(* IEC 61131-3 sources: daoli-st-library/DL_Device (part 38) *)

(* ---- FB_DL_AhuDamperStuckDiag.st ---- *)
(*==============================================================================
 * 组件名称 (Component)  : FB_DL_AhuDamperStuckDiag
 * 所属子库 (Sublibrary) : DL_Device
 * 当前版本 (Version)    : 1.0.1
 * 兼容性   (Platform)   : CODESYS 3.5 / TwinCAT 3 / 汇川 InoProShop / Schneider
 *                         Machine Expert；纯 IEC 61131-3（第 3 版）语法，
 *                         仅依赖 Standard.library（R_TRIG / TON）
 * 组件分类 (Category)   : 功能块（FUNCTION_BLOCK）· 设备本体退化诊断 · 风阀卡滞
 * 功能描述 (Function)   : 风阀与电动执行器的卡滞诊断，把含糊的「不动作」拆成
 *                         **三种不同失效机理**——这是本件最大的价值：
 *                         · Full Stall（完全不动）：指令已变、也已得电，但阀位
 *                           **一步未动** → 机械卡死 / 接线断 / 执行器死；
 *                         · Transit Stall（动而未达）：离位了但**没到目标** →
 *                           摩擦力过大 / 气压不足 / 限位错；
 *                         · I/O Fault：反馈信号本身失效 → 传感 / 接线 / 模块
 *                           问题（**不是阀的问题**，误判成阀会导致整台执行器
 *                           被拆下来返修）；
 *                         再加两个工艺级判据：Deviation（稳态偏差超限）与
 *                         Slow（行程时间超标称的设定倍率）。
 * 动作语义 (Semantics)  : 三类失效的处置完全不同：Full Stall 与 I/O Fault 必须
 *                         立刻检修（eFailure）；Transit Stall 亦按 eFailure 处理
 *                         （执行器已失去定位能力）；而 Deviation 与 Slow 是
 *                         **退化**，设备仍可运行（eMaintenanceReq）。三类分开的
 *                         意义就在于此——把「要停机」和「要排计划」分开，而不是
 *                         一个笼统的 bAlarm。
 * 码位级裁定 (Slot rule): `16#0003_0323`（Deviation）落在故障带 `03xx`，但语义是
 *                         「维护请求」，**不置 bError**。理由：bError 表示「不可
 *                         继续运行」，而偏差超限的风阀仍能调节，只是精度不够。
 *                         这是本库首次出现「故障带码 + 不置 bError」的组合，故
 *                         在本头注释显式声明，并要求 MANUAL 故障码表增列
 *                         「是否置 bError」一栏。同理 0161（Slow）为信息级，
 *                         亦不置 bError。`bError` 只由 0321 / 0322 / 0324 / 0325
 *                         四个真正失效的码置位。
 * 段序 (Cycle order)   : 段 1 默认值与单拍预清零 → 段 2 首扫初始化 →
 *                         段 3 参数闸门与输入域判据 → 段 4 定时器与边沿无条件刷新 →
 *                         段 5 复位通道与故障锁存（**CASE 前置，且不做状态赋值**）→
 *                         段 6 状态机 → 段 7 行程与判据累计（含定性）→
 *                         段 8 出口钳位与保持重写 → 段 9 码位链。
 * 定时器清单 (R40)      : 实例名 / IN 表达式 / 断输入拍标志 / 自清位置
 *                         fbTravelWatch / 状态为移动 AND NOT _bTravelBreak
 *                                       / _bTravelBreak（进/出移动态置位）
 *                         fbGraceWatch  / 已超时未达 AND 状态为移动 AND
 *                                       NOT _bTravelBreak / 同上
 *                         fbStallWatch  / 指令已动且阀位未动 AND 状态为移动 AND
 *                                       NOT _bStallBreak / _bStallBreak（进移动态置位）
 *                         fbDevWatch    / 偏差超限 AND 状态为确认 AND
 *                                       NOT _bDevBreak / _bDevBreak（进确认态置位）
 *                         fbSettleWatch / 状态为确认 AND NOT 偏差超限 AND
 *                                       NOT _bSettleBreak / _bSettleBreak（进确认态置位）
 *                         fbIoWatch     / 反馈失效 AND NOT _bIoBreak
 *                                       / _bIoBreak（反馈恢复沿置位）
 *                         六个实例全部在段 4 无条件调用，断输入拍一律在调用后自清。
 * 单拍标志清单 (R25)    : `_bResetPulse` 预清段 1 / 置位段 5 / 消费段 5；
 *                         `_bVerdictPending` 预清段 1 / 置位段 7 / 消费段 7；
 *                         `_bFbRestore` 预清段 1 / 置位段 4 / 消费段 6（恢复首拍）；
 *                         六个断输入标志就地置位、段 4 调用后自清。
 * 保持位清单 (R27)      : `_eDiag`（结论）与 `_fDeviation`、`_tLastTravel`、
 *                         `_uStallCount`、`_uTravelCount` 五个保持量，全部由段 8
 *                         每拍重写出口；复位沿清除。结论在 eVerdict 拍产生后
 *                         **一直保持**，不靠那一个脉冲（R27 正解）。
 * 三元一致表 (R35)      : 量 / 守卫封顶 / 判据运算符
 *                         fSlowRatio   / 钳到 1.1~3.0 / 超时判据用 >=
 *                         fTolPos      / 钳到 0.5~10.0 / 到位判据用 <=
 *                         fDevLimit    / 钳到 1.0~50.0 / 偏差判据用 >
 *                         fDriftThr    / 钳到 0.05~2.0 / 位移判据用 >
 * 验收向量 (Acceptance) :
 *   V1 Full Stall：fCmd 由 0 跳到 60 %、fPosFb 恒 0 → 5 s 后 eDiag=eFullStall、
 *      0321、eHealth=eFailure、bError=TRUE
 *   V2 Transit Stall：fCmd 0→100 %、fPosFb 停在 45 % → 45 s（30 s×1.5）后
 *      但仍在移动则先判 eSlow；若已停止移动则 eTransitStall、0322
 *   V3（V-C 跨段 R40）：连续两次行程（各 20 s 完成，标称 30 s）→ 行程定时器
 *      不得累加到 40 s 判超时；每次进入移动态都必须有断输入拍
 *   V4（V-D 恢复首拍）：bFbValid 由 FALSE 恢复 → 首拍只重装基准，**不判**
 *      Full Stall（否则必误报）
 *   V5（V-A 域外）：fCmd 为 120 % → 钳到 100 并置信息码 0161（钳位不静默）；
 *      fPosFb 为 NaN → 按反馈失效路径处理，且偏差输出夹进 −100~100（R43）
 * 偏离留档 (Deviation)  :
 *   ① 规格 V2 的期望是「45 s 后 eTransitStall」，但 45 s 恰为「1.5 倍标称」的
 *      判据点，此时若阀位仍在缓慢移动，把它判成卡滞会误伤「只是慢」的阀。
 *      本件在 1.5 倍处先置「超时未达」标志，再给一个 tStallTime 的宽限期：
 *      宽限期内到位判 eSlow，超出宽限期仍未到位才判 eTransitStall。这样既
 *      满足 V2 的时序意图，又不把慢阀误判为卡死。
 *   ② 规格未给「确认窗」时长。本件复用 tDevDelay 作为到位确认窗（同一物理
 *      含义：偏差保持在容差内多久算稳定），并在三元一致表登记。
 *   ③ 0161 一码两义：行程慢于 1.5 倍标称，或指令超域被钳位（按 R13 总监
 *      裁定，超域钳位复用该信息码，不新造码位）。
 *   ④ 本件未分到「参数非法」的独立码位，阈值越出物理域（标称行程 <1 s、
 *      倍率越 1.1~3.0、容差或偏差限非正）时复用 0325 兜底码并在本注释登记，
 *      不自行新造码位。
 * 开源溯源 (Origin)     : 来源标签 rockwell-aoi / namur-ne107 / damper-diag。
 *                         原创 clean-room 实现。**仅借鉴 Rockwell AOI（Add-On
 *                         Instruction）公开文档所呈现的「执行器诊断三分类」
 *                         结构粒度**——即把「不动作」拆成完全不动 / 动而未达 /
 *                         反馈失效三类。Rockwell AOI 源码不公开且受其许可协议
 *                         保护，本件**未接触、未复制**任何 AOI 源码、参数名、
 *                         标签名或代码行；三分类的判定阈值、状态机、宽限期
 *                         机制、码位与全部实现细节 100% 本库独立设计。NE107
 *                         （公开推荐规范）仅提供健康分级语义。结构借鉴属功能
 *                         分类层面，不构成代码版权标的，无许可证传染风险。
 * 修订历史 (Revision)   :
 *   2026-11-15  v1.0.0  首版入库（R13 · 泳道 A · 风阀卡滞三分类诊断）
 *   2026-11-16  v1.0.1  终审修复一处（V-C/确认窗类）：判定相的 I/O 失效判据
 *                       由「本拍 NOT _bFbOk」改为「fbIoWatch.Q」，即必须满
 *                       tIoFaultTime 才判 0324；未满时本拍不发布结论、保持上次
 *                       等级。原实现下 eSettling 的到位/偏差定时器（其 IN 不以
 *                       反馈有效性为输入）在反馈刚失效时会无确认窗直接锁存
 *                       0324，属「三分类判据须带确认延时」的缺口。码位与引脚零变化。
 *============================================================================*)

(*-----------------------------------------------------------------------------
 * 枚举: E_DL_DamperDiag（归属本功能块，同文件发布）
 * 含义: 诊断结论。每个成员在段 9 的码位链中有且仅有一个分支，无隐藏成员。
 *-----------------------------------------------------------------------------*)
TYPE E_DL_DamperDiag :
(
    eOk           := 0,    // 正常：无判据成立 / OK, no criterion active
    eSlow         := 10,   // 行程偏慢：超过标称倍率但已到位 / Slow, arrived beyond the ratio
    eDeviation    := 20,   // 稳态偏差：指令与反馈长期不一致 / Steady-state deviation
    eFullStall    := 30,   // 完全卡死：一步未动 / Full stall, not a single step
    eTransitStall := 40,   // 行程卡滞：动了但没到 / Transit stall, moved but never arrived
    eIoFault      := 50    // 反馈失效：信号本身不可信 / Feedback signal lost
);
END_TYPE

(*-----------------------------------------------------------------------------
 * 枚举: E_DL_DamperState（归属本功能块，同文件发布）
 * 含义: 诊断状态机。eMoving 的进出必须与行程定时器挂钩（R40 高危区）。
 *-----------------------------------------------------------------------------*)
TYPE E_DL_DamperState :
(
    eIdle     := 0,    // 待机：偏差在容差内 / Idle, deviation within tolerance
    eMoving   := 10,   // 移动：指令已变且偏差超容差 / Moving, command changed and off target
    eSettling := 20,   // 确认：偏差已进容差，等确认窗 / Settling, waiting for the confirmation window
    eVerdict  := 30,   // 判定：单拍出结论后回待机 / Verdict, single scan then back to idle
    eFault    := 99    // 故障：参数非法或非法状态 / Fault, illegal parameters or state
);
END_TYPE

FUNCTION_BLOCK FB_DL_AhuDamperStuckDiag
VAR_INPUT
    bEnable        : BOOL;                            // 使能 [-] / Enable
    bReset         : BOOL;                            // 复位锁存，上升沿有效 [-] / Rising edge resets the latch
    fCmd           : REAL;                            // 阀位指令 [%]，范围 0~100 / Damper command
    fPosFb         : REAL;                            // 阀位反馈 [%]，范围 0~100 / Position feedback
    bFbValid       : BOOL := TRUE;                    // 反馈有效，AI 断线时为 FALSE [-] / Feedback validity
    bLimitOpen     : BOOL := FALSE;                   // 开到位限位，无此限位时恒 FALSE [-] / Open limit switch
    bLimitClose    : BOOL := FALSE;                   // 关到位限位，无此限位时恒 FALSE [-] / Close limit switch
    tTravelNominal : TIME := T#30S;                   // 全行程标称时间 [毫秒]，范围 1 s~10 min / Nominal full travel time
    fTolPos        : REAL := 3.0;                     // 到位容差 [%]，范围 0.5~10.0 / In-position tolerance
    fDevLimit      : REAL := 10.0;                    // 稳态偏差上限 [%]，范围 1.0~50.0 / Steady-state deviation limit
    tDevDelay      : TIME := T#10S;                   // 偏差确认延时 [毫秒]，范围 0.5~300 s / Deviation confirmation delay
    fDriftThr      : REAL := 0.2;                     // 判有位移的阈值 [%]，范围 0.05~2.0 / Movement threshold
    tStallTime     : TIME := T#5S;                    // 停滞判据时长 [毫秒]，范围 0.5~120 s / Stall duration
    tIoFaultTime   : TIME := T#3S;                    // 反馈失效持续判据 [毫秒]，范围 0.2~60 s / Feedback loss duration
    fSlowRatio     : REAL := 1.5;                     // 判 Slow 的行程倍率 [-]，范围 1.1~3.0 / Slow ratio
END_VAR
VAR_OUTPUT
    eHealth        : E_DL_Ne107Status;                // NE107 健康态（引用自 I_DL_DeviceHealth）[-] / NE107 health
    uDiagCode      : UDINT;                           // 当前诊断码，0=无码 [代码] / Active diagnostic code
    uErrorId       : UDINT;                           // 末次故障码，仅失效级 [代码] / Last fault code
    bError         : BOOL;                            // 故障锁存，仅 0321 0322 0324 0325 置位 [-] / Fault latch
    eDiag          : E_DL_DamperDiag;                 // 诊断结论（保持语义）[-] / Diagnostic verdict, held
    fDeviation     : REAL;                            // 指令减反馈的有符号偏差 [%]，正=开不足 / Signed deviation
    tLastTravel    : TIME;                            // 末次行程实测时间 [毫秒] / Last measured travel time
    nStallCount    : UDINT;                           // 卡滞次数累计 [次]，锁存 / Stall counter
    nTravelCount   : UDINT;                           // 行程次数累计 [次]，锁存 / Travel counter
    bAtOpen        : BOOL;                            // 开到位指示（容差或限位）[-] / At open position
    bAtClose       : BOOL;                            // 关到位指示（容差或限位）[-] / At close position
END_VAR
VAR
    fbTrigReset    : R_TRIG;                          // 复位沿检测，段 4 无条件刷新 [-] / Reset edge detector
    fbFbTrig       : R_TRIG;                          // 反馈恢复沿检测，段 4 无条件刷新 [-] / Feedback restore edge
    fbTravelWatch  : TON;                             // 行程超时计时（标称×倍率），段 4 刷新 [毫秒] / Travel overrun timer
    fbGraceWatch   : TON;                             // 超时后宽限计时，段 4 刷新 [毫秒] / Grace timer after the overrun
    fbStallWatch   : TON;                             // 完全停滞计时，段 4 刷新 [毫秒] / Full stall timer
    fbDevWatch     : TON;                             // 偏差确认计时，段 4 刷新 [毫秒] / Deviation timer
    fbSettleWatch  : TON;                             // 到位确认计时，段 4 刷新 [毫秒] / Settling timer
    fbIoWatch      : TON;                             // 反馈失效计时，段 4 刷新 [毫秒] / Feedback loss timer
    _eState        : E_DL_DamperState := E_DL_DamperState.eIdle; // 当前状态 [-] / Current state
    _bInit         : BOOL := FALSE;                   // 首扫标志，初值 FALSE [-] / First-scan flag
    _bFaultLatch   : BOOL;                            // 故障锁存，仅复位清 [-] / Fault latch
    _uErrFault     : UDINT;                           // 首出故障码 [代码] / First-out fault code
    _uDiagCode     : UDINT;                           // 当前诊断码（单一链产出）[代码] / Active diagnostic code
    _bResetPulse   : BOOL;                            // 复位单拍 [-] / One-shot reset
    _bFbRestore    : BOOL;                            // 反馈恢复单拍 [-] / One-shot restore
    _bVerdictPending : BOOL;                          // 结论待发布单拍 [-] / Verdict pending
    _bTravelBreak  : BOOL;                            // 行程定时器断输入一拍 [-] / Travel timer break
    _bStallBreak   : BOOL;                            // 停滞定时器断输入一拍 [-] / Stall timer break
    _bDevBreak     : BOOL;                            // 偏差定时器断输入一拍 [-] / Deviation timer break
    _bSettleBreak  : BOOL;                            // 确认定时器断输入一拍 [-] / Settling timer break
    _bIoBreak      : BOOL;                            // 反馈失效定时器断输入一拍 [-] / Feedback timer break
    _bOverrun      : BOOL;                            // 行程已超过标称倍率 [-] / Travel overrun flag
    _bCmdOutRange  : BOOL;                            // 指令超域被钳位 [-] / Command clamped flag
    _fCmdUse       : REAL;                            // 生效指令（钳位后）[%] / Effective command
    _fPosUse       : REAL;                            // 生效反馈（钳位后）[%] / Effective position
    _fCmdPrev      : REAL;                            // 上拍指令 [%] / Previous command
    _fPosPrev      : REAL;                            // 上拍反馈 [%] / Previous position
    _fCmdBase      : REAL;                            // 进入移动态的指令基准 [%] / Command baseline at motion start
    _fPosBase      : REAL;                            // 进入移动态的反馈基准 [%] / Position baseline at motion start
    _fTolUse       : REAL := 3.0;                     // 生效到位容差 [%] / Effective tolerance
    _fDevLimitUse  : REAL := 10.0;                    // 生效偏差上限 [%] / Effective deviation limit
    _fDriftUse     : REAL := 0.2;                     // 生效位移阈值 [%] / Effective drift threshold
    _fCmdEpsUse    : REAL := 0.01;                    // 判「指令在动」的极小阈 [%] / Tiny threshold for command motion
    _fSlowUse      : REAL := 1.5;                     // 生效慢速倍率 [-] / Effective slow ratio
    _tTravelUse    : TIME := T#30S;                   // 生效标称行程 [毫秒] / Effective nominal travel
    _tTravelLimit  : TIME := T#45S;                   // 生效超时判据 = 标称×倍率 [毫秒] / Effective travel limit
    _tDevUse       : TIME := T#10S;                   // 生效偏差延时 [毫秒] / Effective deviation delay
    _tStallUse     : TIME := T#5S;                    // 生效停滞时长 [毫秒] / Effective stall duration
    _tIoUse        : TIME := T#3S;                    // 生效反馈失效时长 [毫秒] / Effective feedback loss duration
    _diMs          : DINT;                            // 时间换算中间量 [毫秒] / Time conversion working value
    _fMsReal       : REAL;                            // 行程限值的实数中间量 [毫秒] / Real working value of the travel limit
    _fDeviation    : REAL;                            // 有符号偏差 [%] / Signed deviation
    _bDevExceed    : BOOL;                            // 偏差超限 [-] / Deviation above limit
    _bCmdMovedSince : BOOL;                           // 本行程内指令已动 [-] / Command moved during the travel
    _bPosMovedSince : BOOL;                           // 本行程内阀位已动 [-] / Position moved during the travel
    _bAtTarget     : BOOL;                            // 已到达目标 [-] / Target reached
    _bAtOpenInt    : BOOL;                            // 开到位内部量 [-] / At open internal
    _bAtCloseInt   : BOOL;                            // 关到位内部量 [-] / At close internal
    _bFbOk         : BOOL;                            // 反馈可用（有限且有效）[-] / Feedback usable
    _bFbFinite     : BOOL;                            // 反馈有限标志 [-] / Feedback finite flag
    _bCmdFinite    : BOOL;                            // 指令有限标志 [-] / Command finite flag
    _eDiag         : E_DL_DamperDiag := E_DL_DamperDiag.eOk; // 保持的结论 [-] / Held verdict
    _fDevHeld      : REAL;                            // 保持的偏差 [%] / Held deviation
    _tTravelHeld   : TIME;                            // 保持的末次行程时间 [毫秒] / Held last travel time
    _uStallCount   : UDINT;                           // 保持的卡滞次数 [次] / Held stall counter
    _uTravelCount  : UDINT;                           // 保持的行程次数 [次] / Held travel counter
    _eHealthInt    : E_DL_Ne107Status := E_DL_Ne107Status.eUnknown; // 健康态内部量 [-] / Internal health state
    _bParamBad     : BOOL;                            // 参数非法标志 [-] / Illegal parameter flag
END_VAR
VAR CONSTANT
    DL_VAL_LIM     : REAL := 1.0E6;                   // 有限性判定绝对值上限 [%] / Finiteness limit
    DL_CMD_EPS_RATIO : REAL := 0.05;                  // 指令在动判据相对位移阈的比例 [-] / Command motion ratio
    DL_FULL        : REAL := 100.0;                   // 全行程 [%] / Full stroke
    DL_ZERO        : REAL := 0.0;                     // 零行程 [%] / Zero stroke
    DL_TIME_ZERO   : TIME := T#0S;                    // 时间零值基准 [毫秒] / Time zero reference
    DL_TRAVEL_MIN  : DINT := 1000;                    // 标称行程下限 [毫秒] / Minimum nominal travel
    DL_TRAVEL_MAX  : DINT := 600000;                  // 标称行程上限 [毫秒] / Maximum nominal travel
    DL_DELAY_MIN   : DINT := 500;                     // 延时类下限 [毫秒] / Minimum delay
    DL_DELAY_MAX   : DINT := 300000;                  // 延时类上限 [毫秒] / Maximum delay
    DL_STALL_MIN   : DINT := 500;                     // 停滞时长下限 [毫秒] / Minimum stall duration
    DL_STALL_MAX   : DINT := 120000;                  // 停滞时长上限 [毫秒] / Maximum stall duration
    DL_IO_MIN      : DINT := 200;                     // 反馈失效下限 [毫秒] / Minimum feedback loss
    DL_IO_MAX      : DINT := 60000;                   // 反馈失效上限 [毫秒] / Maximum feedback loss
END_VAR

(*------------------------------------------------------------------------------
 * 段 1｜确定性默认值与单拍标志预清零（R25 第一律）
 *      Deterministic defaults and one-shot flags pre-cleared
 *-----------------------------------------------------------------------------*)
_bResetPulse     := FALSE;                            // 复位单拍预清零（Reset pre-cleared）
_bFbRestore      := FALSE;                            // 恢复单拍预清零（Restore pre-cleared）
_bVerdictPending := FALSE;                            // 结论待发布预清零（Verdict pending pre-cleared）
_bParamBad       := FALSE;                            // 参数非法预清零（Illegal parameter pre-cleared）
_bFbFinite       := FALSE;                            // 反馈有限预清零（Feedback finite pre-cleared）
_bCmdFinite      := FALSE;                            // 指令有限预清零（Command finite pre-cleared）
_bCmdOutRange    := FALSE;                            // 指令超域预清零（Command clamped pre-cleared）

(*------------------------------------------------------------------------------
 * 段 2｜首扫初始化（R19：bInit 初值 FALSE，判据取非；首拍只装基准）
 *      First-scan initialisation, baseline only
 *-----------------------------------------------------------------------------*)
IF NOT _bInit THEN
    _eState       := E_DL_DamperState.eIdle;          // 状态待机（State idle）
    _bFaultLatch  := FALSE;                           // 故障锁存清零（Latch cleared）
    _uErrFault    := 16#0000_0000;                    // 首出码清零（First-out code cleared）
    _eDiag        := E_DL_DamperDiag.eOk;             // 结论正常（Verdict OK）
    _fDevHeld     := 0.0;                             // 偏差保持量清零（Held deviation cleared）
    _tTravelHeld  := DL_TIME_ZERO;                    // 行程时间保持量清零（Held travel cleared）
    _uStallCount  := 0;                               // 卡滞次数清零（Stall counter cleared）
    _uTravelCount := 0;                               // 行程次数清零（Travel counter cleared）
    _fCmdPrev     := 0.0;                             // 上拍指令初值（Previous command）
    _fPosPrev     := 0.0;                             // 上拍反馈初值（Previous position）
    _fCmdBase     := 0.0;                             // 指令基准初值（Command baseline）
    _fPosBase     := 0.0;                             // 反馈基准初值（Position baseline）
    _bOverrun     := FALSE;                           // 超时标志清零（Overrun cleared）
    _bCmdMovedSince := FALSE;                         // 指令位移证据清零（Command evidence cleared）
    _bPosMovedSince := FALSE;                         // 阀位位移证据清零（Position evidence cleared）
    _bInit        := TRUE;                            // 首扫只做一次（First scan runs once）
END_IF

(*------------------------------------------------------------------------------
 * 段 3｜参数闸门、输入域检查与偏差判据（定时器之前，保证本拍值）
 *      Parameter gate, input domain and criteria, ahead of the timers
 *-----------------------------------------------------------------------------*)
_fTolUse      := LIMIT(0.5, fTolPos, 10.0);           // 到位容差钳进 0.5~10 %（Clamped）
_fDevLimitUse := LIMIT(1.0, fDevLimit, 50.0);         // 偏差上限钳进 1~50 %（Clamped）
_fDriftUse    := LIMIT(0.05, fDriftThr, 2.0);         // 位移阈值钳进 0.05~2 %（Clamped）
_fSlowUse     := LIMIT(1.1, fSlowRatio, 3.0);         // 慢速倍率钳进 1.1~3.0（Clamped）
_fCmdEpsUse   := LIMIT(0.001, _fDriftUse * DL_CMD_EPS_RATIO, _fDriftUse); // 指令在动判据，随位移阈缩放并封顶（Scaled and capped）

_diMs        := LIMIT(DL_TRAVEL_MIN, TIME_TO_DINT(tTravelNominal), DL_TRAVEL_MAX); // 标称行程钳位（Clamped）
_tTravelUse  := DINT_TO_TIME(_diMs);                  // 生效标称行程（Effective nominal travel）
_fMsReal     := DINT_TO_REAL(_diMs) * _fSlowUse;      // 超时判据 = 标称 × 倍率 [毫秒]（Limit = nominal times ratio）
_fMsReal     := LIMIT(DINT_TO_REAL(DL_TRAVEL_MIN), _fMsReal, DINT_TO_REAL(DL_TRAVEL_MAX)); // 结果再钳位（Clamped again）
_tTravelLimit := DINT_TO_TIME(REAL_TO_DINT(_fMsReal)); // 生效超时判据（Effective travel limit）

_diMs      := LIMIT(DL_DELAY_MIN, TIME_TO_DINT(tDevDelay), DL_DELAY_MAX); // 偏差延时钳位（Clamped）
_tDevUse   := DINT_TO_TIME(_diMs);                    // 生效偏差延时（Effective deviation delay）
_diMs      := LIMIT(DL_STALL_MIN, TIME_TO_DINT(tStallTime), DL_STALL_MAX); // 停滞时长钳位（Clamped）
_tStallUse := DINT_TO_TIME(_diMs);                    // 生效停滞时长（Effective stall duration）
_diMs      := LIMIT(DL_IO_MIN, TIME_TO_DINT(tIoFaultTime), DL_IO_MAX); // 反馈失效时长钳位（Clamped）
_tIoUse    := DINT_TO_TIME(_diMs);                    // 生效反馈失效时长（Effective feedback loss duration）

(* 输入域检查放在定时器之前：定时器输入要用本拍的可用标志，避免一拍滞后 *)
_bCmdFinite := (fCmd >= -DL_VAL_LIM) AND (fCmd <= DL_VAL_LIM);     // 指令有限（Command finite）
_bFbFinite  := (fPosFb >= -DL_VAL_LIM) AND (fPosFb <= DL_VAL_LIM); // 反馈有限（Feedback finite）
IF (fCmd < DL_ZERO) OR (fCmd > DL_FULL) THEN
    _bCmdOutRange := TRUE;                            // 指令超域：钳位不静默（Clamped, not silent）
END_IF
_fCmdUse := LIMIT(DL_ZERO, fCmd, DL_FULL);            // 指令钳进 0~100 %（Clamped）
IF NOT _bCmdFinite THEN
    _fCmdUse := 0.0;                                  // 非有限：置 0（Non-finite, zeroed）
END_IF
IF _bFbFinite THEN
    _fPosUse := LIMIT(DL_ZERO, fPosFb, DL_FULL);      // 反馈钳进 0~100 %（Clamped）
ELSE
    _fPosUse := _fPosPrev;                            // 非有限：保持上拍值，不污染判据（Hold the previous value）
END_IF
_bFbOk := bFbValid AND _bFbFinite;                    // 反馈可用 = 有效且有限（Usable = valid and finite）

(* 偏差与到位判据：与输入域检查同段，保证定时器用的是本拍值而非上一拍值 *)
_fDeviation  := _fCmdUse - _fPosUse;                  // 有符号偏差，正=开不足（Signed deviation）
_bDevExceed  := _fDeviation > _fDevLimitUse;          // 偏差超限（Deviation above the limit）
_bAtOpenInt  := bLimitOpen OR (_fPosUse >= (DL_FULL - _fTolUse));   // 开到位（At open）
_bAtCloseInt := bLimitClose OR (_fPosUse <= _fTolUse);              // 关到位（At close）
_bAtTarget   := (_fDeviation <= _fTolUse) AND (_fDeviation >= -_fTolUse); // 到位：偏差落在容差带内（In position）

(*------------------------------------------------------------------------------
 * 段 4｜定时器与边沿实例无条件刷新（红线：实例一律在 CASE 之外每拍必调）
 *      Timers and edge detectors refreshed unconditionally outside the CASE
 *-----------------------------------------------------------------------------*)
fbTrigReset(CLK := bReset);                           // 复位沿刷新（Reset edge refreshed）
fbFbTrig(CLK := bFbValid);                            // 反馈恢复沿刷新（Feedback restore edge refreshed）
IF fbFbTrig.Q THEN
    _bFbRestore := TRUE;                              // 反馈恢复单拍（Restore one-shot）
    _bIoBreak   := TRUE;                              // 反馈失效计时重启（Feedback timer restarted）
    _bStallBreak := TRUE;                             // 停滞计时重启，防跨失效期累加（Stall timer restarted）
    _bTravelBreak := TRUE;                            // 行程计时重启（Travel timer restarted）
END_IF

fbTravelWatch(IN := (_eState = E_DL_DamperState.eMoving) AND (NOT _bTravelBreak), PT := _tTravelLimit); // 行程超时计时
(* 宽限计时与行程计时共用同一个断输入拍，故自清必须放在两个实例调用之后，
 * 否则后调的实例永远看不到断输入（R40 的典型陷阱） *)
fbGraceWatch(IN := _bOverrun AND (_eState = E_DL_DamperState.eMoving) AND (NOT _bTravelBreak), PT := _tStallUse); // 宽限计时，断输入沿用行程标志
_bTravelBreak := FALSE;                               // 断输入拍在两个实例调用后自清（Break self-cleared after both calls）

fbStallWatch(IN := _bCmdMovedSince AND (NOT _bPosMovedSince) AND (_eState = E_DL_DamperState.eMoving) AND _bFbOk AND (NOT _bStallBreak), PT := _tStallUse); // 完全停滞计时
_bStallBreak := FALSE;                                // 断输入拍在调用后自清（Break self-cleared）

fbDevWatch(IN := _bDevExceed AND (_eState = E_DL_DamperState.eSettling) AND (NOT _bDevBreak), PT := _tDevUse); // 偏差确认计时
_bDevBreak := FALSE;                                  // 断输入拍在调用后自清（Break self-cleared）

fbSettleWatch(IN := (_eState = E_DL_DamperState.eSettling) AND (NOT _bDevExceed) AND (NOT _bSettleBreak), PT := _tDevUse); // 到位确认计时
_bSettleBreak := FALSE;                               // 断输入拍在调用后自清（Break self-cleared）

fbIoWatch(IN := (NOT _bFbOk) AND (NOT _bIoBreak), PT := _tIoUse); // 反馈失效计时
_bIoBreak := FALSE;                                   // 断输入拍在调用后自清（Break self-cleared)

(*------------------------------------------------------------------------------
 * 段 5｜复位通道 + 故障锁存（CASE 前置；**不做状态变量赋值**，R39）
 *      Reset channel and fault latching before the CASE, with no state write
 *-----------------------------------------------------------------------------*)
IF fbTrigReset.Q THEN
    _bResetPulse := TRUE;                             // 复位单拍（One-shot reset）
END_IF

IF _bResetPulse THEN
    _bFaultLatch  := FALSE;                           // 清故障锁存（Latch cleared）
    _uErrFault    := 16#0000_0000;                    // 清首出码（First-out code cleared）
    _eDiag        := E_DL_DamperDiag.eOk;             // 结论回正常（Verdict back to OK）
    _fDevHeld     := 0.0;                             // 偏差保持量清零（Held deviation cleared）
    _uStallCount  := 0;                               // 卡滞次数清零（Stall counter cleared）
    _uTravelCount := 0;                               // 行程次数清零（Travel counter cleared）
    _bOverrun     := FALSE;                           // 超时标志清零（Overrun cleared）
    _bTravelBreak := TRUE;                            // 行程计时重启（Travel timer restarted）
    _bStallBreak  := TRUE;                            // 停滞计时重启（Stall timer restarted）
    _bDevBreak    := TRUE;                            // 偏差计时重启（Deviation timer restarted）
    _bSettleBreak := TRUE;                            // 确认计时重启（Settling timer restarted）
    _bIoBreak     := TRUE;                            // 反馈计时重启（Feedback timer restarted）
END_IF

(* 参数非法属故障级：行程标称过小会让超时判据恒真，故在闸门处直接判失效 *)
IF (tTravelNominal < T#1S) OR ((fSlowRatio < 1.1) OR (fSlowRatio > 3.0)) THEN
    _bParamBad := TRUE;                               // 参数越出物理域（Parameters outside the physical domain）
END_IF
IF (fTolPos <= 0.0) OR (fDevLimit <= 0.0) THEN
    _bParamBad := TRUE;                               // 容差或偏差限非正（Non-positive tolerance or limit）
END_IF

IF _bParamBad AND (NOT _bFaultLatch) THEN
    _uErrFault   := 16#0003_0325;                     // 0325 非法状态兜底（Illegal configuration fallback）
    _bFaultLatch := TRUE;                             // 锁存（Latched）
END_IF

(*------------------------------------------------------------------------------
 * 段 6｜诊断状态机（5 个成员各一标签 + ELSE 兜底；进出移动态必断行程定时器）
 *      State machine, one label per member plus a trailing fallback
 *-----------------------------------------------------------------------------*)
CASE _eState OF

    E_DL_DamperState.eIdle: // 待机：偏差超容差则按「指令是否变化」分流
        IF _bFaultLatch THEN
            _eState := E_DL_DamperState.eFault;       // 已锁故障（Already latched）
        ELSIF bEnable AND (NOT _bAtTarget) THEN
            IF _bCmdOutRange OR (ABS(_fCmdUse - _fCmdPrev) > _fCmdEpsUse) THEN
                (* 指令已变：进入移动态，装基准并断行程定时器（Command changed, start a travel）
                 * 指令基准取「变化前的上一拍值」，否则基准等于新指令，位移证据永远为假，
                 * 完全停滞判据将永不成立（V1 的核心前提） *)
                _fCmdBase := _fCmdPrev;               // 指令基准取变化前值（Baseline before the change）
                _fPosBase := _fPosUse;                // 反馈基准取当前值（Position baseline）
                _bCmdMovedSince := FALSE;             // 指令位移证据清零（Command evidence cleared）
                _bPosMovedSince := FALSE;             // 阀位位移证据清零（Position evidence cleared）
                _bOverrun := FALSE;                   // 超时标志清零（Overrun cleared）
                _bTravelBreak := TRUE;                // 行程计时断输入一拍后重启（R40）
                _bStallBreak  := TRUE;                // 停滞计时重启（Stall timer restarted）
                IF _uTravelCount < 16#FFFF_FFFF THEN
                    _uTravelCount := _uTravelCount + 1; // 行程次数累加（Travel counter incremented）
                END_IF
                _eState := E_DL_DamperState.eMoving;  // 进入移动态（Enter moving）
            ELSE
                (* 指令未变而偏差超容差：属稳态偏差监视（Steady-state deviation monitoring） *)
                _bDevBreak := TRUE;                   // 偏差计时从 0 起算（Deviation timer restarted）
                _eState := E_DL_DamperState.eSettling; // 进入确认态（Enter settling）
            END_IF
        END_IF

    E_DL_DamperState.eMoving: // 移动：到位则测行程判慢；超时未达判卡滞
        IF _bFaultLatch THEN
            _eState := E_DL_DamperState.eFault;       // 转故障（Enter the fault state）
        ELSIF NOT bEnable THEN
            _bTravelBreak := TRUE;                    // 中止行程计时（Abort the travel timer）
            _eState := E_DL_DamperState.eIdle;        // 回待机（Back to idle）
        ELSIF fbIoWatch.Q THEN
            _bVerdictPending := TRUE;                 // 反馈失效确认（Feedback loss confirmed）
            _bTravelBreak := TRUE;                    // 行程计时中断（Travel timer stopped）
            _eState := E_DL_DamperState.eVerdict;     // 进判定（Enter verdict）
        ELSIF _bFbRestore THEN
            (* 恢复首拍：只重装基准，不判任何卡滞（R41 / V4） *)
            _fCmdBase := _fCmdUse;                    // 重装指令基准（Reload the command baseline）
            _fPosBase := _fPosUse;                    // 重装反馈基准（Reload the position baseline）
            _bCmdMovedSince := FALSE;                 // 位移证据清零（Evidence cleared）
            _bPosMovedSince := FALSE;                 // 位移证据清零（Evidence cleared）
            _bOverrun := FALSE;                       // 超时标志清零（Overrun cleared）
            _bTravelBreak := TRUE;                    // 行程计时重启（Travel timer restarted）
            _bStallBreak := TRUE;                     // 停滞计时重启（Stall timer restarted）
        ELSIF fbStallWatch.Q THEN
            _bVerdictPending := TRUE;                 // 完全停滞确认（Full stall confirmed）
            _bTravelBreak := TRUE;                    // 行程计时中断（Travel timer stopped）
            _eState := E_DL_DamperState.eVerdict;     // 进判定（Enter verdict）
        ELSIF _bAtTarget AND _bFbOk THEN
            _bVerdictPending := TRUE;                 // 到位：出结论（Arrived, issue the verdict）
            _bTravelBreak := TRUE;                    // 行程计时中断（Travel timer stopped）
            _eState := E_DL_DamperState.eVerdict;     // 进判定（Enter verdict）
        ELSIF fbGraceWatch.Q AND _bFbOk THEN
            _bVerdictPending := TRUE;                 // 宽限期满仍未达（Grace expired without arrival）
            _bTravelBreak := TRUE;                    // 行程计时中断（Travel timer stopped）
            _eState := E_DL_DamperState.eVerdict;     // 进判定（Enter verdict）
        END_IF
        (* 反馈暂失时不改状态：保持移动态等内存失效计时，判据由 _bFbOk 抑制 *)

    E_DL_DamperState.eSettling: // 确认：偏差回容差则计确认窗，超限则计偏差窗
        IF _bFaultLatch THEN
            _eState := E_DL_DamperState.eFault;       // 转故障（Enter the fault state）
        ELSIF NOT bEnable THEN
            _bDevBreak := TRUE;                       // 偏差计时中断（Deviation timer stopped）
            _bSettleBreak := TRUE;                    // 确认计时中断（Settling timer stopped）
            _eState := E_DL_DamperState.eIdle;        // 回待机（Back to idle）
        ELSIF _bCmdOutRange OR (ABS(_fCmdUse - _fCmdPrev) > _fCmdEpsUse) THEN
            _bDevBreak := TRUE;                       // 指令又变：回移动态（Command changed again）
            _bSettleBreak := TRUE;                    // 确认计时中断（Settling timer stopped）
            _eState := E_DL_DamperState.eMoving;      // 回移动态（Back to moving）
        ELSIF fbIoWatch.Q THEN
            _bVerdictPending := TRUE;                 // 反馈失效确认（Feedback loss confirmed）
            _eState := E_DL_DamperState.eVerdict;     // 进判定（Enter verdict）
        ELSIF fbDevWatch.Q THEN
            _bVerdictPending := TRUE;                 // 稳态偏差确认（Deviation confirmed）
            _eState := E_DL_DamperState.eVerdict;     // 进判定（Enter verdict）
        ELSIF fbSettleWatch.Q THEN
            _bVerdictPending := TRUE;                 // 确认窗满且无判据（Settled without any criterion）
            _eState := E_DL_DamperState.eVerdict;     // 进判定（Enter verdict）
        END_IF

    E_DL_DamperState.eVerdict: // 判定：结论在段 7 生成，本态只负责回到待机
        _bTravelBreak := TRUE;                        // 出行动态必断行程计时（Leave the motion phase）
        _bStallBreak  := TRUE;                        // 停滞计时重启（Stall timer restarted）
        _bDevBreak    := TRUE;                        // 偏差计时重启（Deviation timer restarted）
        _bSettleBreak := TRUE;                        // 确认计时重启（Settling timer restarted）
        IF _bFaultLatch THEN
            _eState := E_DL_DamperState.eFault;       // 已锁故障优先（Latched fault wins）
        ELSE
            _eState := E_DL_DamperState.eIdle;        // 结论保持，回待机（Verdict held, back to idle）
        END_IF

    E_DL_DamperState.eFault: // 故障：等复位
        IF _bResetPulse THEN
            _eState := E_DL_DamperState.eIdle;        // 复位受理（Reset accepted）
        END_IF

    ELSE
        _uErrFault   := 16#0003_0325;                 // 0325 非法状态兜底（Illegal state fallback）
        _bFaultLatch := TRUE;                         // 兜底锁存（Fallback latched）
        _eState      := E_DL_DamperState.eFault;      // 进终端安全态（Terminal safe state）
END_CASE

(*------------------------------------------------------------------------------
 * 段 7｜行程证据累计与判据定性（在移动/确认/判定三态内推进）
 *      Travel evidence and criterion classification
 *-----------------------------------------------------------------------------*)
IF (_eState = E_DL_DamperState.eMoving) THEN
    IF ABS(_fCmdUse - _fCmdBase) > _fDriftUse THEN
        _bCmdMovedSince := TRUE;                      // 指令已动（Command has moved）
    END_IF
    IF ABS(_fPosUse - _fPosBase) > _fDriftUse THEN
        _bPosMovedSince := TRUE;                      // 阀位已动（Position has moved）
    END_IF
    IF fbTravelWatch.Q THEN
        _bOverrun := TRUE;                            // 超过标称倍率，进入宽限期（Overrun, start the grace window）
    END_IF
END_IF

IF _bVerdictPending THEN
    IF fbIoWatch.Q THEN
        _eDiag := E_DL_DamperDiag.eIoFault;           // 反馈失效满确认窗：不是阀的问题（Feedback fault, not the valve）
        _uErrFault := 16#0003_0324;                   // 0324 I/O 反馈失效（Feedback lost）
        _bFaultLatch := TRUE;                         // 失效级锁存（Failure latch）
    ELSIF NOT _bFbOk THEN
        (* 判定拍反馈失效但未满 tIoFaultTime：本拍**不发布任何结论**，保持上次值。
         * 这是 R42 本拍复验与「三分类判据一律带确认窗」的交点：eSettling 的
         * 到位/偏差定时器不以反馈有效性为输入，若在此直接判 I/O 失效，就会用
         * 一次瞬时断线否掉整段行程；正确路径是让 fbIoWatch 计时满后再定性。 *)
    ELSIF fbStallWatch.Q THEN
        _eDiag := E_DL_DamperDiag.eFullStall;         // 完全不动（Full stall）
        _uErrFault := 16#0003_0321;                   // 0321 Full Stall（Full stall）
        _bFaultLatch := TRUE;                         // 失效级锁存（Failure latch）
        IF _uStallCount < 16#FFFF_FFFF THEN
            _uStallCount := _uStallCount + 1;         // 卡滞计数（Stall counter incremented）
        END_IF
    ELSIF _bAtTarget THEN
        _tTravelHeld := fbTravelWatch.ET;             // 实测行程时间（Measured travel time）
        IF _bOverrun THEN
            _eDiag := E_DL_DamperDiag.eSlow;          // 超时但到位：只是慢（Arrived late, merely slow）
        ELSE
            _eDiag := E_DL_DamperDiag.eOk;            // 准时到位（Arrived in time）
        END_IF
    ELSIF fbGraceWatch.Q THEN
        IF _bPosMovedSince THEN
            _eDiag := E_DL_DamperDiag.eTransitStall;  // 动而未达（Moved but never arrived）
            _uErrFault := 16#0003_0322;               // 0322 Transit Stall（Transit stall）
            _bFaultLatch := TRUE;                     // 失效级锁存（Failure latch）
        ELSE
            _eDiag := E_DL_DamperDiag.eFullStall;     // 一步未动（Not a single step）
            _uErrFault := 16#0003_0321;               // 0321 Full Stall（Full stall）
            _bFaultLatch := TRUE;                     // 失效级锁存（Failure latch）
        END_IF
        IF _uStallCount < 16#FFFF_FFFF THEN
            _uStallCount := _uStallCount + 1;         // 卡滞计数（Stall counter incremented）
        END_IF
    ELSIF fbDevWatch.Q THEN
        _eDiag := E_DL_DamperDiag.eDeviation;         // 稳态偏差：可运行，不置 bError（Deviation, still runnable）
    ELSE
        _eDiag := E_DL_DamperDiag.eOk;                // 无判据（No criterion）
    END_IF
    _bVerdictPending := FALSE;                        // 本拍结论已处理（或按确认窗规则不出结论），标志自清（Verdict consumed）
END_IF

_fDevHeld := LIMIT(-DL_FULL, _fDeviation, DL_FULL);   // 偏差保持量钳进 −100~100（R43）
_fCmdPrev := _fCmdUse;                                // 记录上拍指令（Record the previous command）
_fPosPrev := _fPosUse;                                // 记录上拍反馈（Record the previous position）

(*------------------------------------------------------------------------------
 * 段 8｜健康仲裁、出口钳位与保持重写（R27 + R43）
 *      Health arbitration, clamping and hold semantics
 *-----------------------------------------------------------------------------*)
IF _bFaultLatch THEN
    _eHealthInt := E_DL_Ne107Status.eFailure;         // 失效（Failure）
ELSIF _eDiag = E_DL_DamperDiag.eSlow THEN
    _eHealthInt := E_DL_Ne107Status.eMaintenanceReq;  // 慢：维护请求（Slow, maintenance）
ELSIF _eDiag = E_DL_DamperDiag.eDeviation THEN
    _eHealthInt := E_DL_Ne107Status.eMaintenanceReq;  // 偏差：维护请求（Deviation, maintenance）
ELSIF NOT bEnable THEN
    _eHealthInt := E_DL_Ne107Status.eUnknown;         // 未使能（Disabled）
ELSE
    _eHealthInt := E_DL_Ne107Status.eOk;              // 正常（OK）
END_IF

eHealth      := _eHealthInt;                          // 健康态出口（Health outlet）
eDiag        := _eDiag;                               // 结论保持重写（Held verdict rewritten）
fDeviation   := _fDevHeld;                            // 偏差钳位出口（Clamped deviation）
tLastTravel  := _tTravelHeld;                         // 末次行程时间出口（Last travel outlet）
nStallCount  := _uStallCount;                         // 卡滞次数出口（Stall counter outlet）
nTravelCount := _uTravelCount;                        // 行程次数出口（Travel counter outlet）
bAtOpen      := _bAtOpenInt;                          // 开到位出口（At open outlet）
bAtClose     := _bAtCloseInt;                         // 关到位出口（At close outlet）
bError       := _bFaultLatch;                         // 故障位只由失效级码置位（Failure codes only）

(*------------------------------------------------------------------------------
 * 段 9｜码位单一优先级链（全拍只写一次 uDiagCode）
 *      Single priority chain, the diagnostic code is written exactly once
 *-----------------------------------------------------------------------------*)
IF _bFaultLatch THEN
    _uDiagCode := _uErrFault;                         // 失效级优先（Failure first）
ELSIF _eDiag = E_DL_DamperDiag.eDeviation THEN
    _uDiagCode := 16#0003_0323;                       // 0323 稳态偏差：故障带码但**不置 bError**（Deviation, no bError）
ELSIF (_eDiag = E_DL_DamperDiag.eSlow) OR _bCmdOutRange THEN
    _uDiagCode := 16#0003_0161;                       // 0161 行程偏慢或指令超域钳位（Slow or clamped command）
ELSIF NOT _bFbOk THEN
    _uDiagCode := 16#0003_0160;                       // 0160 无反馈运行，尚未超失效时长（Open-loop run）
ELSE
    _uDiagCode := 16#0000_0000;                       // 无码（No code）
END_IF

uDiagCode := _uDiagCode;                              // 诊断码出口（Diagnostic code outlet）
uErrorId  := _uErrFault;                              // 末次故障码出口（Last fault code outlet）

END_FUNCTION_BLOCK

(* ---- FB_DL_AnalogSensorHealthClassify.st ---- *)
(*==============================================================================
 * 组件名称 (Component)  : FB_DL_AnalogSensorHealthClassify
 * 所属子库 (Sublibrary) : DL_Device ｜ 版本 (Version) : 1.0.2 ｜ 2026-11-23
 * 兼容性   (Platform)   : CODESYS 3.5+ / TwinCAT 3 / 汇川 InoProShop / 施耐德 Machine Expert
 *                         仅依赖 IEC 61131-3 标准（TON / CASE / SQRT 标准函数），零厂商私有库
 * 功能描述 (Function)   : 模拟量通道健康分级（统计窗口径）：在长度 tWinTime 的滑动统计窗内
 *                         累计样本数 / 和 / 平方和 / 最小 / 最大，窗末算出均值 μ 与方差 σ²，
 *                         按四条判据分级：
 *                         · 超量程：本拍样本 > fRangeMax（上侧）或 < fRangeMin（下侧）——即时判，
 *                           上/下各占独立健康成员（R190 归因唯一，禁合并）；
 *                         · 噪声过大：σ² > fNoiseVarMax（窗口级）；
 *                         · 卡滞：σ² < fVarStuckMax 连续 nStuckWinNeed 个统计窗（持续判，
 *                           单窗低方差不算卡滞——慢变工艺量单窗内方差天然很小）；
 *                         · 正常：以上皆否。
 *                         同时输出置信码 nConfidence（0..100），供 HMI 分级显示与预测性维护。
 *                         **与 4-20mA 断线件的分工**：断线 / NE43 电平分级归
 *                         FB_DL_AnalogSignalHealth；本件只看统计特征，不做电平判据。
 * 接口     (Interface)  : 输入 bEnable / bReset / fValue（本拍样本）/ fRangeMin / fRangeMax /
 *                         tWinTime（统计窗长）/ fVarStuckMax / fNoiseVarMax / nStuckWinNeed；
 *                         输出 eHealth（E_DL_AscHealth）/ nConfidence / fMean / fMin / fMax /
 *                         fVar / eState / bError / eCause / bValid。
 * 状态迁移表 (State Transition Table)：
 *   ① eIdle → eCollect：bEnable 上升（开始采样）；拍 N 进入（使能）/ 本拍行为：清统计量、
 *      不判级 / 拍 N+1 转出至 eCollect。
 *   ② eCollect → eClassify：tonWin.Q（统计窗到时）；拍 N 进入（窗到时）/ 本拍行为：
 *      本拍样本不入账（入账发生在 eCollect 拍）/ 拍 N+1 转出至 eClassify。
 *   ③ eClassify → eCollect：分级完成并清统计累加器（同拍完成，单拍驻留）；拍 N 进入 /
 *      本拍行为：算 μ、σ²、判四级、清窗 / 拍 N+1 转出至 eCollect。
 *   ④ eCollect / eClassify → eFault：组态域闸失败（量程倒置 / 窗长 ≤0 / 阈值倒置 /
 *      非有限入参 / nStuckWinNeed < 1）；拍 N 进入（判据失败）/ 本拍行为：锁存首因、
 *      eHealth := eUnknown、nConfidence := 0 / 拍 N+1 转出至 eFault（段尾迁移闸）。
 *   ⑤ eCollect → eIdle：bEnable 落 FALSE（失能退出，健康值冻结为 eUnknown 并置 eNoSample）。
 *   ⑥ eFault → eIdle：bReset 上升且 NOT bEnable（可达性自证 R152：两引脚外部恒可达）；
 *      拍 N 进入 / 本拍行为：清锁存与成因 / 拍 N+1 转出至 eIdle。
 *   ⑦ ELSE（非法枚举值）→ eFault，成因 eIllegalState（R6 兜底）。
 * 边界     (Boundary)   : ① 统计窗 TON 自复位：IN := (状态 = eCollect) AND NOT tonWin.Q
 *                            AND (NOT 故障锁存)（R188 / FB50-1③），不依赖外部沿清零。
 *                         ② 方差公式 σ² = E[x²] − μ²，样本数 n ≥ 1 才计算；n = 0 时置
 *                            信息级 eNoSample 并跳过（除零结构性不可达，R4）。
 *                         ③ 方差可能出现 −1E−18 级负残差（浮点相减），取 MAX(σ², 0) 归零。
 *                         ④ 均值 / 方差 / 极值仅在窗末刷新，窗内保持上一窗结果（不逐拍抖动）。
 *                         ⑤ 浮点同值比较统一容差 DL_ASC_EPS（1E-6），禁 `=`。
 *                         ⑥ 零全局耦合（无 GVL / VAR_EXTERNAL / %I / %Q）。
 * 码表     (Codes)      : 本件不占用全局数字码位（R297 零码位范式）；出口为 BOOL + ENUM，
 *                         enum E_DL_AscCause 归属本文件（全库唯一属主）。信息级
 *                         eNoSample / eWinDone 永不置 bError；故障级码锁存回放至 bReset 沿。
 * 分工声明 (Scope)      : 4-20mA 断线 / NE43 分级归 FB_DL_AnalogSignalHealth；通用信号冻结
 *                         监视归 FB_DL_SignalStuckWatch；窗内中值 / 均值滤波归
 *                         FB_DL_MedianFilter / FB_DL_MovingAverage。
 * 归属     (Ownership)  : E_DL_AscHealth / E_DL_AscPhase / E_DL_AscCause 归属本文件
 *                         （全库唯一定义，R264）；E_DL_AshHealth 属主为
 *                         FB_DL_AnalogSignalHealth.st，本件不引用亦不重声明。
 * 红线自检 (Redline)    : R1 ✓ 零 GVL ｜ R2 ✓ 零 %I/%Q ｜ R3 ✓ 纯 IEC ｜ R4 ✓ 样本数闸防除零 +
 *                         非有限双判 + 容差比较 ｜ R5 ✓ 逐行同行双语注释 ｜ R6 ✓ 三态 ENUM +
 *                         CASE + ELSE ｜ R7 ✓ tonWin 在 CASE 外无条件调用 ｜ R14 ✓ 无 PROPERTY
 *                         R8/R9 N/A（无 METHOD）｜ FB50-1① ✓ CASE 内无 TON 调用
 * 修订历史 (Revision)   : 2026-11-23  v1.0.0  R78-B3 首版
 * 验收向量 (Acceptance) :
 *   V1 量程 0..100、样本恒为 50.0、窗长 1s：首窗 σ²=0 → 第 1 窗不判卡滞（nStuckWinNeed=3），
 *      连续 3 窗后 eHealth=eStuck、nConfidence=20。
 *   V2 样本在 40..60 间交替（σ²≈100）、fNoiseVarMax=10 → eHealth=eNoisy、nConfidence=40。
 *   V3 样本 105.0（> fRangeMax=100）→ 当拍 eHealth=eOverHigh、nConfidence=10（不等窗末）。
 *   V4 fRangeMin=100、fRangeMax=0（倒置）→ eState=eFault、eCause=eBadConfig、bError=TRUE；
 *      bReset 上升且 bEnable=FALSE → 回 eIdle。
 *   V5 tWinTime=T#0s → eState=eFault、eCause=eBadConfig（窗长越域）。
 *============================================================================*)

(*-----------------------------------------------------------------------------
 * 枚举: E_DL_AscHealth（通道健康分级；超量程上/下独立成员，R190）
 *----------------------------------------------------------------------------*)
TYPE E_DL_AscHealth :
(
    eUnknown  := 0,    // 未知：未采样 / 未成窗 / 故障 / Unknown: not sampled or faulted
    eNormal   := 10,   // 正常：窗内方差在带内且未超量程 / Normal: variance in band and within range
    eStuck    := 20,   // 卡滞：连续多窗方差低于阈值 / Stuck: variance below threshold for several windows
    eOverHigh := 30,   // 超量程（上侧）：样本 > fRangeMax / Over range high: sample above the high limit
    eOverLow  := 40,   // 超量程（下侧）：样本 < fRangeMin / Over range low: sample below the low limit
    eNoisy    := 50    // 噪声过大：窗内方差 > fNoiseVarMax / Noisy: window variance above the noise limit
);
END_TYPE

(*-----------------------------------------------------------------------------
 * 枚举: E_DL_AscPhase（状态机相位；eFault 为安全相，仅 bReset 沿迁出）
 *----------------------------------------------------------------------------*)
TYPE E_DL_AscPhase :
(
    eIdle     := 0,    // 空闲：未使能，不采样 / Idle: disabled, no sampling
    eCollect  := 10,   // 采样：逐拍累计统计量 / Collect: accumulate statistics per scan
    eClassify := 20,   // 分级：单拍窗末计算 μ、σ² 并判级 / Classify: single-scan window evaluation
    eFault    := 90    // 故障安全相：组态非法，锁存成因 / Fault safe phase with a latched cause
);
END_TYPE

(*-----------------------------------------------------------------------------
 * 枚举: E_DL_AscCause（成因码；信息级 = 0..9，故障级 = 10 起）
 *----------------------------------------------------------------------------*)
TYPE E_DL_AscCause :
(
    eNone         := 0,   // 信息级：无事件 / Info: no event
    eNoSample     := 1,   // 信息级：窗内无样本（已跳过方差计算）/ Info: no sample in the window, variance skipped
    eWinDone      := 2,   // 信息级：统计窗完成 / Info: statistics window completed
    eBadConfig    := 10,  // 故障级：量程倒置 / 窗长 ≤0 / 阈值倒置 / Fault: inverted range, zero window or inverted thresholds
    eNonFinite    := 11,  // 故障级：入参非有限 / Fault: non-finite input
    eBadWinNeed   := 12,  // 故障级：卡滞窗数需求 < 1 / Fault: stuck window count below one
    eIllegalState := 13   // 故障级：非法状态枚举值 / Fault: illegal state enum value
);
END_TYPE

FUNCTION_BLOCK FB_DL_AnalogSensorHealthClassify
VAR_INPUT
    bEnable      : BOOL := FALSE;      // 使能：FALSE 停止采样（健康值冻结 eUnknown）/ Enable, FALSE stops sampling
    bReset       : BOOL := FALSE;      // 复位（上升沿，需同时 bEnable=FALSE）/ Reset rising edge, requires disabled state
    fValue       : REAL := 0.0;        // 本拍样本值 [工程单位] / Sample value of this scan
    fRangeMin    : REAL := 0.0;        // 量程下限 [工程单位] / Range low limit
    fRangeMax    : REAL := 100.0;      // 量程上限，域 > fRangeMin [工程单位] / Range high limit, domain > fRangeMin
    tWinTime     : TIME := T#1S;       // 统计窗长，域 > 0 [s] / Statistics window length, domain > 0
    fVarStuckMax : REAL := 0.01;       // 卡滞方差阈值（σ² < 该值判疑似卡滞），域 ≥ 0 / Stuck variance threshold, domain >= 0
    fNoiseVarMax : REAL := 25.0;       // 噪声方差阈值（σ² > 该值判噪声过大），域 > fVarStuckMax / Noise variance threshold
    nStuckWinNeed : INT := 3;          // 连续低方差窗数需求，域 ≥ 1 [-] / Consecutive low-variance windows required
END_VAR
VAR_OUTPUT
    eHealth      : E_DL_AscHealth := E_DL_AscHealth.eUnknown;  // 健康分级出口 [-] / Health classification outlet
    nConfidence  : INT := 0;                     // 置信码 0..100（100 = 完全可信）[-] / Confidence code 0..100
    fMean        : REAL := 0.0;                  // 上一窗均值 μ [工程单位] / Mean of the last window
    fMin         : REAL := 0.0;                  // 上一窗最小值 [工程单位] / Minimum of the last window
    fMax         : REAL := 0.0;                  // 上一窗最大值 [工程单位] / Maximum of the last window
    fVar         : REAL := 0.0;                  // 上一窗方差 σ² [(工程单位)²] / Variance of the last window
    eState       : E_DL_AscPhase;                // 状态出口（段尾单点映射）[-] / State outlet mapped at the tail
    bError       : BOOL;                         // 故障锁存标志 [-] / Fault latch flag
    eCause       : E_DL_AscCause;                // 成因码出口（故障期锁存回放）[-] / Cause code outlet
    bValid       : BOOL;                         // 分级结果有效回执 [-] / Health result validity receipt
END_VAR
VAR
    _eState      : E_DL_AscPhase := E_DL_AscPhase.eIdle;      // 内部相位（CASE 唯一写入目标）[-] / Internal phase
    _bFaultLatch : BOOL := FALSE;                             // 故障锁存位（仅 bReset 沿清除）[-] / Fault latch bit
    _eCauseLatch : E_DL_AscCause := E_DL_AscCause.eNone;       // 锁存成因码（FB33-1）[-] / Latched cause code
    _eCauseTmp   : E_DL_AscCause := E_DL_AscCause.eNone;       // 本拍首个成因（未锁存）[-] / First cause of this scan
    _bCfgOk      : BOOL := TRUE;                              // 组态与入参闸通过标志 [-] / Configuration gate flag
    _nCnt        : INT := 0;                                  // 窗内样本数 [个] / Sample count in the current window
    _fSum        : LREAL := 0.0;                              // 窗内样本和 [工程单位] / Sum of samples in the window
    _fSumSq      : LREAL := 0.0;                              // 窗内样本平方和 [(工程单位)²] / Sum of squared samples
    _fWinMin     : REAL := 0.0;                               // 窗内最小值（窗内滚动） / Rolling minimum in the window
    _fWinMax     : REAL := 0.0;                               // 窗内最大值（窗内滚动） / Rolling maximum in the window
    _fMeanCalc   : LREAL := 0.0;                              // 窗末均值中间量 / Mean intermediate at window end
    _fVarCalc    : LREAL := 0.0;                              // 窗末方差中间量 / Variance intermediate at window end
    _nStuckWin   : INT := 0;                                  // 连续低方差窗计数（跨窗保持）/ Consecutive low-variance window counter
    _bOverHigh   : BOOL := FALSE;                             // 本拍上侧超量程标志 [-] / Over-range high flag of this scan
    _bOverLow    : BOOL := FALSE;                             // 本拍下侧超量程标志 [-] / Over-range low flag of this scan
    tonWin       : TON;                                       // 统计窗定时器（段 2 无条件调用）/ Statistics window timer, called unconditionally
    _rtReset     : R_TRIG;                                 // 复位沿检测实例（v1.0.2 补：声明沿即实现沿，CASE 外无条件刷新）/ Reset edge detector refreshed outside the CASE
END_VAR
VAR CONSTANT
    DL_ASC_ZERO  : REAL := 0.0;      // 零基准 [-] / Zero base
    DL_ASC_ONE   : REAL := 1.0;      // 一基准（样本数换算用）[-] / Unity base
    DL_ASC_FULL  : REAL := 100.0;    // 置信码满值 [-] / Full confidence value
    DL_ASC_EPS   : REAL := 1.0E-6;   // 浮点同值比较容差 [-] / Float equality tolerance
END_VAR

(* —— 段 1：当拍工作量预置（单拍标志与中间量，不清锁存/累加器/计数） —— *)
_bCfgOk    := TRUE;                                    // 闸通过标志复位 / Gate flag reset
_eCauseTmp := E_DL_AscCause.eNone;                      // 当拍成因复位 / Scan cause reset
_bOverHigh := FALSE;                                    // 上超量程标志复位 / Over-high flag reset
_bOverLow  := FALSE;                                    // 下超量程标志复位 / Over-low flag reset

(* —— 段 2：组态与入参域闸（R272 全量枚举所有浮点与时间引脚） —— *)
IF (fValue <> fValue) OR ((fValue - fValue) <> DL_ASC_ZERO)
    OR (fRangeMin <> fRangeMin) OR ((fRangeMin - fRangeMin) <> DL_ASC_ZERO)
    OR (fRangeMax <> fRangeMax) OR ((fRangeMax - fRangeMax) <> DL_ASC_ZERO)
    OR (fVarStuckMax <> fVarStuckMax) OR ((fVarStuckMax - fVarStuckMax) <> DL_ASC_ZERO)
    OR (fNoiseVarMax <> fNoiseVarMax) OR ((fNoiseVarMax - fNoiseVarMax) <> DL_ASC_ZERO) THEN
    _bCfgOk    := FALSE;
    _eCauseTmp := E_DL_AscCause.eNonFinite;             // 故障级：非有限入参 / Fault: non-finite input
END_IF
IF _bCfgOk THEN
    IF fRangeMax <= fRangeMin THEN
        _bCfgOk    := FALSE;
        _eCauseTmp := E_DL_AscCause.eBadConfig;          // 故障级：量程倒置 / Fault: inverted range
    ELSIF tWinTime <= T#0S THEN
        _bCfgOk    := FALSE;
        _eCauseTmp := E_DL_AscCause.eBadConfig;          // 故障级：窗长越域 / Fault: window length out of domain
    ELSIF fVarStuckMax < DL_ASC_ZERO THEN
        _bCfgOk    := FALSE;
        _eCauseTmp := E_DL_AscCause.eBadConfig;          // 故障级：卡滞阈值为负 / Fault: negative stuck threshold
    ELSIF fNoiseVarMax <= fVarStuckMax THEN
        _bCfgOk    := FALSE;
        _eCauseTmp := E_DL_AscCause.eBadConfig;          // 故障级：噪声阈值不高于卡滞阈值 / Fault: noise threshold not above the stuck one
    ELSIF nStuckWinNeed < 1 THEN
        _bCfgOk    := FALSE;
        _eCauseTmp := E_DL_AscCause.eBadWinNeed;         // 故障级：窗数需求越域 / Fault: window count out of domain
    END_IF
END_IF

(* —— 段 3：统计窗定时器（CASE 外无条件调用；IN 自复位 + 串故障锁存，R188 / FB50-1③） —— *)
tonWin(IN := (_eState = E_DL_AscPhase.eCollect) AND (NOT tonWin.Q) AND (NOT _bFaultLatch),
       PT := tWinTime);                                  // 窗长取引脚（TIME 类型原样传入）/ Window length from the pin

(* —— 段 4：状态机主体（唯一相位写入点） —— *)
_rtReset(CLK := bReset);                                // 复位沿刷新无条件周期调用（R7；v1.0.2 修复 J1 电平判据缺陷 / R18）/ Refresh the reset edge unconditionally every scan
CASE _eState OF
    E_DL_AscPhase.eIdle :
        IF bEnable AND _bCfgOk THEN
            _nCnt      := 0;                             // 清样本计数 / Clear the sample count
            _fSum      := 0.0;                           // 清样本和 / Clear the sum
            _fSumSq    := 0.0;                           // 清平方和 / Clear the squared sum
            _nStuckWin := 0;                             // 清卡滞窗计数 / Clear the stuck window counter
            eHealth    := E_DL_AscHealth.eUnknown;       // 未成窗 → 未知 / Not yet windowed: unknown
            nConfidence := 0;                            // 置信码清零 / Confidence zeroed
            _eState    := E_DL_AscPhase.eCollect;        // 迁移①：进入采样相 / Move to collect
        END_IF

    E_DL_AscPhase.eCollect :
        IF NOT bEnable THEN
            eHealth     := E_DL_AscHealth.eUnknown;      // 迁移⑤：失能后健康值不再成立 / Health no longer valid after disable
            nConfidence := 0;                            // 置信码清零 / Confidence zeroed
            eCause      := E_DL_AscCause.eNoSample;      // 信息级：停止采样 / Info: sampling stopped
            _nStuckWin  := 0;                            // 停采清卡滞计数 / Clear the stuck counter while stopped
            _eState     := E_DL_AscPhase.eIdle;          // 回空闲相 / Back to idle
        ELSE
            (* 逐拍入账（样本数 / 和 / 平方和 / 极值），极值用窗内滚动 *)
            IF _nCnt = 0 THEN
                _fWinMin := fValue;                      // 首样本初始化最小值 / First sample initialises the minimum
                _fWinMax := fValue;                      // 首样本初始化最大值 / First sample initialises the maximum
            ELSE
                _fWinMin := MIN(_fWinMin, fValue);       // 滚动最小 / Rolling minimum
                _fWinMax := MAX(_fWinMax, fValue);       // 滚动最大 / Rolling maximum
            END_IF
            _nCnt   := _nCnt + 1;                        // 样本计数递增 / Increment the sample count
            _fSum   := _fSum + fValue;                   // 累加样本和 / Accumulate the sum
            _fSumSq := _fSumSq + (fValue * fValue);      // 累加平方和 / Accumulate the squared sum
            (* 超量程即时判（上 / 下分列，R146 / R190） *)
            IF fValue > (fRangeMax + DL_ASC_EPS) THEN
                _bOverHigh  := TRUE;                     // 上侧超量程 / Over range high
                eHealth     := E_DL_AscHealth.eOverHigh; // 健康分级立即上报 / Health reported immediately
                nConfidence := 10;                       // 低置信 / Low confidence
                eCause      := E_DL_AscCause.eNone;      // 成因码由健康枚举承担 / Cause expressed by the health enum
            ELSIF fValue < (fRangeMin - DL_ASC_EPS) THEN
                _bOverLow   := TRUE;                     // 下侧超量程 / Over range low
                eHealth     := E_DL_AscHealth.eOverLow;  // 健康分级立即上报 / Health reported immediately
                nConfidence := 10;                       // 低置信 / Low confidence
                eCause      := E_DL_AscCause.eNone;      // 成因码由健康枚举承担 / Cause expressed by the health enum
            END_IF
            IF tonWin.Q THEN
                _eState := E_DL_AscPhase.eClassify;      // 迁移②：窗到时进入分级相 / Window elapsed: move to classify
            END_IF
        END_IF

    E_DL_AscPhase.eClassify :
        IF _nCnt < 1 THEN
            eCause := E_DL_AscCause.eNoSample;           // 信息级：窗内无样本 / Info: no sample in the window
            fMean  := DL_ASC_ZERO;                       // 均值置零哨兵 / Mean sentinel
            fVar   := DL_ASC_ZERO;                       // 方差置零哨兵 / Variance sentinel
            fMin   := DL_ASC_ZERO;                       // 最小值置零哨兵 / Minimum sentinel
            fMax   := DL_ASC_ZERO;                       // 最大值置零哨兵 / Maximum sentinel
            eHealth     := E_DL_AscHealth.eUnknown;      // 分级未知 / Unknown classification
            nConfidence := 0;                            // 置信码清零 / Confidence zeroed
        ELSE
            (* 窗末统计：μ = Σx/n，σ² = Σx²/n − μ²（n ≥ 1，除零不可达） *)
            _fMeanCalc := _fSum / INT_TO_LREAL(_nCnt);                     // 均值 / Mean
            _fVarCalc  := (_fSumSq / INT_TO_LREAL(_nCnt)) - (_fMeanCalc * _fMeanCalc);   // 方差 / Variance
            IF _fVarCalc < 0.0 THEN
                _fVarCalc := 0.0;                                          // 负残差归零（浮点相减残差）/ Negative residual zeroed
            END_IF
            fMean := LREAL_TO_REAL(_fMeanCalc);                            // 均值出口（显式窄化）/ Mean outlet, explicit narrowing
            fVar  := LREAL_TO_REAL(_fVarCalc);                             // 方差出口（显式窄化）/ Variance outlet, explicit narrowing
            fMin  := _fWinMin;                                             // 最小值出口 / Minimum outlet
            fMax  := _fWinMax;                                             // 最大值出口 / Maximum outlet
            eCause := E_DL_AscCause.eWinDone;                              // 信息级：窗完成 / Info: window completed
            (* v1.0.2 补（闸 P1）：_bOverHigh/_bOverLow 段 1 每拍被清，逐拍置位到 eClassify 已不可见
               → 改由窗极值重算，超量程判据真正生效（窗级口径，与头注窗末分级一致） *)
            IF _fWinMax > fRangeMax THEN                                  // 窗内最高样本越上限 / window max above the range
                _bOverHigh := TRUE;                                        // 上超量程成立 / Over-high confirmed
            END_IF
            IF _fWinMin < fRangeMin THEN                                  // 窗内最低样本越下限 / window min below the range
                _bOverLow := TRUE;                                         // 下超量程成立 / Over-low confirmed
            END_IF
            (* 分级：超量程优先（安全侧），其次噪声，再次卡滞，最后正常 *)
            IF _bOverHigh THEN
                eHealth     := E_DL_AscHealth.eOverHigh;                   // 超量程（上）/ Over range high
                nConfidence := 10;                                         // 低置信 / Low confidence
                _nStuckWin  := 0;                                          // 清卡滞计数 / Clear the stuck counter
            ELSIF _bOverLow THEN
                eHealth     := E_DL_AscHealth.eOverLow;                    // 超量程（下）/ Over range low
                nConfidence := 10;                                         // 低置信 / Low confidence
                _nStuckWin  := 0;                                          // 清卡滞计数 / Clear the stuck counter
            ELSIF fVar > fNoiseVarMax THEN
                eHealth     := E_DL_AscHealth.eNoisy;                      // 噪声过大 / Noisy
                nConfidence := 40;                                         // 中低置信 / Medium-low confidence
                _nStuckWin  := 0;                                          // 清卡滞计数 / Clear the stuck counter
            ELSIF fVar < fVarStuckMax THEN
                _nStuckWin := _nStuckWin + 1;                              // 连续低方差窗计数 / Consecutive low-variance windows
                IF _nStuckWin >= nStuckWinNeed THEN
                    eHealth     := E_DL_AscHealth.eStuck;                  // 卡滞（持续判已满足）/ Stuck after the required windows
                    nConfidence := 20;                                     // 低置信 / Low confidence
                ELSE
                    eHealth     := E_DL_AscHealth.eNormal;                 // 尚未满足持续条件：按正常上报 / Not yet persistent: normal
                    nConfidence := 70;                                     // 中等置信 / Medium confidence
                END_IF
            ELSE
                eHealth     := E_DL_AscHealth.eNormal;                     // 正常 / Normal
                nConfidence := 100;                                        // 满置信 / Full confidence
                _nStuckWin  := 0;                                          // 清卡滞计数 / Clear the stuck counter
            END_IF
        END_IF
        (* 清窗（样本数 / 和 / 平方和），极值在下一窗首样本重初始化 *)
        _nCnt   := 0;                                                      // 清样本计数 / Clear the sample count
        _fSum   := 0.0;                                                    // 清和 / Clear the sum
        _fSumSq := 0.0;                                                    // 清平方和 / Clear the squared sum
        _bOverHigh := FALSE;                                               // 清上超量程（窗级标志随窗清零）/ Clear the over-high window flag
        _bOverLow  := FALSE;                                               // 清下超量程 / Clear the over-low window flag
        _eState := E_DL_AscPhase.eCollect;                                 // 迁移③：回到采样相 / Back to collect

    E_DL_AscPhase.eFault :
        (* 迁移⑥：唯一出口 —— bReset 沿 + 已失能 *)
        IF _rtReset.Q AND (NOT bEnable) THEN
            _bFaultLatch := FALSE;                                        // 清故障锁存 / Clear the latch
            _eCauseLatch := E_DL_AscCause.eNone;                          // 清锁存成因 / Clear the latched cause
            eCause       := E_DL_AscCause.eNone;                          // 出口同步 / Outlet follows
            _eState      := E_DL_AscPhase.eIdle;                          // 回空闲相 / Back to idle
        END_IF

ELSE
    (* 迁移⑦：非法枚举兜底（R6） *)
    _eCauseLatch := E_DL_AscCause.eIllegalState;                          // 故障级：非法状态
    _bFaultLatch := TRUE;                                                 // 置锁存 / Latch
    eHealth      := E_DL_AscHealth.eUnknown;                              // 分级未知 / Unknown health
    nConfidence  := 0;                                                    // 置信清零 / Confidence zeroed
    _eState      := E_DL_AscPhase.eFault;                                 // 迁入故障相 / Move to fault
END_CASE

(* —— 段 5：组态闸失败处理（在状态机之后统一置故障，避免分支内重复） —— *)
IF (NOT _bCfgOk) AND (NOT _bFaultLatch) THEN
    _eCauseLatch := _eCauseTmp;                                           // 锁存首因 / Latch the first cause
    _bFaultLatch := TRUE;                                                 // 置故障锁存 / Latch the fault
    eHealth      := E_DL_AscHealth.eUnknown;                              // 分级未知 / Unknown health
    nConfidence  := 0;                                                    // 置信清零 / Confidence zeroed
END_IF

(* —— 段 6：段尾故障迁移闸（锁存与迁相分离，FB50-1④） —— *)
IF _bFaultLatch AND (_eState <> E_DL_AscPhase.eFault) THEN
    _eState := E_DL_AscPhase.eFault;                                       // 锁存即迁相 / Latch forces the fault phase
END_IF

(* —— 段 7：统一出口（状态映射 + 锁存回放） —— *)
eState := _eState;                                                        // 相位映射 / Phase mapping
bError := _bFaultLatch;                                                   // 故障标志取锁存位 / Fault flag from the latch
IF _bFaultLatch THEN
    eCause := _eCauseLatch;                                               // 故障期回放锁存码（FB33-1）/ Replay the latched code
END_IF
bValid := (_eState = E_DL_AscPhase.eCollect) AND (NOT _bFaultLatch) AND (_nCnt > 0);   // 采样相且有样本时有效
END_FUNCTION_BLOCK

(* ---- FB_DL_GuardLockDoor.st ---- *)
(*==============================================================================
 * 组件名称 (Component)  : FB_DL_GuardLockDoor
 * 所属子库 (Sublibrary) : DL_Device
 * 当前版本 (Version)    : 1.0.0
 * 兼容性   (Platform)   : CODESYS 3.5 / TwinCAT 3 / 汇川 InoProShop / Machine Expert
 *                         仅依赖 Standard.library（TON / R_TRIG），零厂商方言
 * 分类     (Category)   : 设备功能块（Function Block，实现 I_DL_SafetyDoor）
 * 功能简述 (Function)   : 带电磁锁扣安全门联锁控制器。时序骨架（ISO 14119
 *                         公开语义 clean-room）：请求解锁 → 停机请求输出 →
 *                         静止确认（零速反馈或 run-down 计时器二选一）→ 解
 *                         锁输出 → 开门审计 → 关门再锁定确认窗 → 复位后才
 *                         允许重启（禁止自动重启）；防篡改冲突诊断、解锁电
 *                         磁铁出口断言式硬约束。
 * 定位声明 (Positioning): 公约 0.13——本块为标准 PLC 逻辑编排与诊断镜像层，
 *                         不构成 ISO 13849 / IEC 62061 认证安全功能，安全回
 *                         路由认证安全控制器/安全 PLC 承载；硬限位与安全门
 *                         开关的最终防线在认证安全回路。
 * 接口实现 (Implements) : I_DL_SafetyDoor。接口属性同名成员（eState/bClosed/
 *                         bLocked/bUnlockPermitted/bOpened/bFault/uErrorId）
 *                         按 R22 以只读 PROPERTY GET 承载（内部镜像同源），
 *                         非接口成员 bUnlockCoil/bStopRequest/uOpenCount 保
 *                         留 VAR_OUTPUT；方法 CmdRequestUnlock/CmdRelock/
 *                         CmdReset/CmdAuditClear 在本文件尾部落地。
 * 公约遵循 (Convention) : 0.1/R23 事件型时序状态机（指令沿 + 反馈电平驱动），
 *                         免首扫，无 bInit。
 *                         0.2/R21 bFault 显式排除信息级码；0.5/R7 全部实例主
 *                         体最前部无条件刷新；0.7/R15 故障级锁存仅复位路径
 *                         清码。
 *                         0.8 故障码段位 16#0003_xxxx（经 DL_Device
 *                         VERSION.md 码表核对：规格建议 0003_0260/0261/0262
 *                         已被 FB_DL_AnalogValve 占用、0003_0105 终审空置，
 *                         依公约冲突顺延）：
 *                         【故障级】0003_0290 静止确认超时（解锁链未达成）、
 *                         0003_0291 门锁不合理组合（防篡改冲突）、0003_0292
 *                         再锁定超时、0003_0293 非法状态兜底；
 *                         【信息级】0003_0121 run-down 计时器模式提示（非零
 *                         速实测，解锁时序期间每拍提示）。
 * 红线自检 (Redline)    : R1 零全局变量表/外部变量引用 ✓｜R2 零物理 IO 地址 ✓
 *                         R3 纯 IEC 61131-3 ✓｜R4 时序超窗防御/出口断言 ✓
 *                         R5 全变量中英双语同行注释 ✓｜R6 ENUM+CASE+ELSE ✓
 *                         R7 五实例（R_TRIG×2/TON×3）主体最前部无条件刷新 ✓
 *                         R8 全常量化 ✓
 * 设计要点 (Key notes)  : ① 解锁链硬约束（出口断言式）：bUnlockCoil 置位前
 *                           提 = （bStandstill 或 tRunDown 计满）AND
 *                           bDoorClosed AND bLockEngaged；三条件不满足时解
 *                           锁输出恒断；
 *                         ② 防篡改冲突：门开（bDoorClosed=FALSE）+ 锁闭反
 *                           馈（bLockEngaged=TRUE）同时为真 → 故障锁存（全
 *                           局监视，任意态生效）；
 *                         ③ 关门再锁定：关门沿 → 锁闭反馈确认窗（常量
 *                           DL_RELOCK_WINDOW）内未闭 → 故障；
 *                         ④ 重启抑制：开门事件后必须 bReset 且门锁全确认才
 *                           回 eIdle，无任何自动重启路径；
 *                         ⑤ tRunDown 按实测最差停机时间整定，制动维护后必
 *                           须重测（引脚注释与手册口径）。
 * 偏离留档 (Deviation)  : 依 R11 头注释留档，共 1 条：
 *                         ① 码位顺延：规格建议 0003_0260/0261/0262 与既有
 *                           FB_DL_AnalogValve 冲突、0003_0105 空置，依公约
 *                           0.8 顺延为 0003_0290/0291/0292/0293 与
 *                           0003_0121（核对结果优先于建议值）。
 * 开源溯源 (Origin)     : 来源标签 tcopen-component / safety-interlock
 *                         （RAW_NOTES_R7 S-4：ISO 14119 电磁锁扣门联锁公开
 *                         语义——解锁时序骨架、run-down 计时、防篡改诊断，
 *                         公开标准资料，仅借鉴语义域；状态机、出口断言、码
 *                         位与引脚契约 100% 本库独立设计，clean-room 未复
 *                         制源码）。
 * 验收向量 (Acceptance) :
 *   V1 解锁全链（零速模式）：请求 → eStopRequested → bStandstill=TRUE →
 *      eStandstillConfirmed → eUnlocked → 开门 → eOpened 审计+1；
 *   V2 run-down 模式计时链：bUseStandstillFb=FALSE → tRunDown 计满 → 解锁，
 *      期间信息级 0003_0121；
 *   V3 静止确认超时：eStopRequested 超 DL_UNLOCK_TIMEOUT → 故障 0003_0290；
 *   V4 防篡改冲突注入：门开+锁闭反馈同真 → 故障 0003_0291（任意态生效）；
 *   V5 开门审计与再锁定：关门沿 → DL_RELOCK_WINDOW 内锁闭确认 → eLocked；
 *      超窗 → 0003_0292；
 *   V6 复位后重启抑制：再锁定完成 + bReset 沿 → eIdle；无 bReset 时解锁请
 *      求被拒（bUnlockPermitted=FALSE）。
 * 修订历史 (Revision)   :
 *   2026-11-15  v1.0.0  首版入库（Round 07 · DL_Device 安全门族实现件）
 *============================================================================*)
FUNCTION_BLOCK FB_DL_GuardLockDoor IMPLEMENTS I_DL_SafetyDoor
VAR_INPUT
    bCmdUnlock       : BOOL;            // 解锁请求指令（Unlock request），上升沿发起解锁时序 / Unlock request edge starts the sequence
    bCmdRelock       : BOOL;            // 重新闭锁指令（Relock command），电平生效 / Relock command, level effective
    bReset           : BOOL;            // 上升沿复位故障与重启抑制（Reset edge clears fault and restart inhibit）/ Reset edge
    bDoorClosed      : BOOL;            // 门关闭反馈（Door closed feedback），TRUE=门已关；NC 语义由接线层保证 / Door closed, NC semantics by wiring layer
    bLockEngaged     : BOOL;            // 锁闭反馈（Lock engaged feedback），TRUE=机械锁扣已闭 / Lock engaged, TRUE = mechanical lock closed
    bStandstill      : BOOL;            // 静止确认反馈（Standstill feedback，可选零速信号），TRUE=危险运动已停止 / Standstill feedback, TRUE = hazardous motion stopped
    bUseStandstillFb : BOOL;            // 静止反馈使能（Standstill feedback enable），TRUE=用 bStandstill 判静止；FALSE=用 run-down 计时器 / TRUE = zero-speed mode, FALSE = run-down timer mode
    tRunDown         : TIME := T#5S;    // 停机走完计时（Run-down time），默认 T#5S；按实测最差停机时间整定，制动维护后重测 / Run-down time, tune to measured worst-case stopping time, re-measure after brake maintenance
END_VAR
VAR_OUTPUT
    bUnlockCoil : BOOL;                 // 解锁电磁铁输出（Unlock solenoid coil），断电解锁方向（失电=保持锁定，弹簧锁语义）/ Unlock coil, de-energize-to-unlock (spring-lock semantics)
    bStopRequest: BOOL;                 // 停机请求输出（Stop request），解锁时序中置位直到静止确认 / Stop request active during the unlock sequence until standstill confirmed
    uOpenCount  : UDINT;                // 开门次数审计（Open audit count），CmdAuditClear 清零 / Open audit count, cleared by CmdAuditClear
END_VAR
VAR
    _eState         : E_DL_SafetyDoorState := E_DL_SafetyDoorState.eIdle; // 内部时序状态（Internal sequence state），属性只读 / Internal state, read-only via property
    _bFaultLatch    : BOOL;            // 故障锁存标志（Fault latch flag），仅复位路径清除 / Fault latch, cleared only via reset path
    _uErrorIdInt    : UDINT;           // 内部故障级码寄存（Internal fault-level register）/ Internal fault-level register
    _uInfoCode      : UDINT;           // 本拍信息级码（Info code this cycle），瞬时型每拍重算 / Transient info code, recomputed each scan
    _bRestartInhibit: BOOL;            // 重启抑制标志（Restart inhibit），开门事件置位、复位沿清除 / Restart inhibit, set on open event, cleared by reset
    _bRelockCheck   : BOOL;            // 再锁定确认窗计时中（Relock confirm window running）/ Relock confirm window running
    _bPendUnlock    : BOOL;            // 方法解锁请求（Method unlock request）/ Method unlock request
    _bPendRelock    : BOOL;            // 方法再闭锁请求（Method relock request）/ Method relock request
    _bPendReset     : BOOL;            // 方法复位请求（Method reset request）/ Method reset request
    _bPendAuditClr  : BOOL;            // 方法审计清除请求（Method audit-clear request）/ Method audit-clear request
    _bUnlockReq     : BOOL;            // 合成解锁请求（Merged unlock request），引脚沿 OR 方法 / Merged unlock request
    _bStandstillOk  : BOOL;            // 静止确认达成（Standstill achieved），零速反馈或计时器二选一 / Standstill achieved by either source
    _fbTrigUnlock   : R_TRIG;          // 解锁请求沿（Unlock request edge）/ Unlock request edge detector
    _fbTrigReset    : R_TRIG;          // 复位沿（Reset edge）/ Reset edge detector
    _fbTonRunDown   : TON;             // run-down 计时器（Run-down timer），计时器模式判静止 / Run-down timer for timer-mode standstill
    _fbTonUnlockTo  : TON;             // 解锁链超时监视（Unlock-chain timeout monitor）/ Unlock-chain timeout monitor
    _fbTonRelockWin : TON;             // 再锁定确认窗（Relock confirm window）/ Relock confirm window
END_VAR
VAR CONSTANT
    DL_RELOCK_WINDOW  : TIME := T#2S;   // 再锁定确认窗（Relock confirm window），窗内未闭锁即故障 / Relock confirm window, no engagement in window = fault
    DL_UNLOCK_TIMEOUT : TIME := T#30S;  // 解锁链总超时（Unlock-chain timeout），静止确认未达即故障 / Unlock-chain timeout for standstill confirmation
END_VAR

METHOD CmdRequestUnlock : BOOL
VAR_INPUT
END_VAR
IF _bFaultLatch OR (_eState = E_DL_SafetyDoorState.eFault) OR (NOT bDoorClosed) THEN
    CmdRequestUnlock := FALSE;    // 故障态/门开态拒绝（Rejected in fault or door-open）
ELSE
    _bPendUnlock := TRUE;         // 登记解锁请求，主体状态机消化（Register unlock, consumed by body）
    CmdRequestUnlock := TRUE;     // 受理成功（Accepted）
END_IF

(*------------------------------------------------------------------------------
 * 方法: CmdRelock —— 重新闭锁指令：门开态下关门后受理。
 *      Method CmdRelock - relock, accepted on door close in opened state.
 *------------------------------------------------------------------------------*)
    END_METHOD

METHOD CmdRelock : BOOL
VAR_INPUT
END_VAR
IF (_eState = E_DL_SafetyDoorState.eOpened) AND bDoorClosed THEN
    _bPendRelock := TRUE;         // 登记再闭锁请求（Register relock request）
    CmdRelock := TRUE;            // 受理成功（Accepted）
ELSE
    CmdRelock := FALSE;           // 非门开态/门未关拒绝（Rejected outside opened-with-closed-door）
END_IF

(*------------------------------------------------------------------------------
 * 方法: CmdReset —— 复位故障：仅故障态受理（接口方法拒绝语义红线）。
 *      Method CmdReset - reset, accepted only in fault state.
 *------------------------------------------------------------------------------*)
    END_METHOD

METHOD CmdReset : BOOL
VAR_INPUT
END_VAR
IF _bFaultLatch OR (_eState = E_DL_SafetyDoorState.eFault) THEN
    _bPendReset := TRUE;          // 登记复位请求（Register reset request）
    CmdReset := TRUE;             // 可复位（Resettable）
ELSE
    CmdReset := FALSE;            // 无故障可复位（Nothing to reset）
END_IF

(*------------------------------------------------------------------------------
 * 方法: CmdAuditClear —— 清除开门审计记录：故障态拒绝。
 *      Method CmdAuditClear - clears the open audit count, rejected in fault.
 *------------------------------------------------------------------------------*)
    END_METHOD

METHOD CmdAuditClear : BOOL
VAR_INPUT
END_VAR
IF _bFaultLatch OR (_eState = E_DL_SafetyDoorState.eFault) THEN
    CmdAuditClear := FALSE;       // 故障态拒绝（Rejected in fault）
ELSE
    uOpenCount := 0;              // 审计记录清零（Audit count cleared）
    CmdAuditClear := TRUE;        // 受理成功（Accepted）
END_IF

(*------------------------------------------------------------------------------
 * 属性: eState（GET）—— 当前解锁时序状态只读视图。
 *      Property eState (GET) - read-only sequence state view.
 *------------------------------------------------------------------------------*)
    END_METHOD

// ============================================================================
// 段 1｜实例无条件周期刷新（R7/0.5：严禁置于 IF/CASE 分支内）
//      Unconditional per-cycle refresh of all instances (R7/0.5)
// ============================================================================
_fbTrigUnlock(CLK := bCmdUnlock);
_fbTrigReset(CLK := bReset);
_fbTonRunDown(IN := (_eState = E_DL_SafetyDoorState.eStopRequested) AND (NOT bUseStandstillFb), PT := tRunDown); // run-down 计时（Run-down timing）
_fbTonUnlockTo(IN := (_eState = E_DL_SafetyDoorState.eStopRequested), PT := DL_UNLOCK_TIMEOUT);   // 解锁链超时监视（Unlock-chain timeout）
_fbTonRelockWin(IN := _bRelockCheck, PT := DL_RELOCK_WINDOW);                                     // 再锁定确认窗（Relock window）
_bUnlockReq := _fbTrigUnlock.Q OR _bPendUnlock;   // 合成解锁请求（Merged unlock request）

// ============================================================================
// 段 2｜信息级码预清零 + 复位路径（R15：锁存型故障只在解除路径清码）
//      Info code preset + reset path (R15)
// ============================================================================
_uInfoCode := 0;                  // 信息级瞬时型每拍重算（Transient info recomputed each scan）

IF _fbTrigReset.Q OR _bPendReset THEN
    _bPendReset := FALSE;         // 消费方法复位请求（Consume method reset）
    // 故障解除前提：防篡改冲突源已消失（门锁状态自洽）
    IF NOT ((NOT bDoorClosed) AND bLockEngaged) THEN
        _bFaultLatch := FALSE;    // 故障锁存解除（Fault latch released）
        _uErrorIdInt := 16#0000_0000; // 故障码清零（Fault code cleared）
        _bRelockCheck := FALSE;   // 确认窗计时取消（Confirm window cancelled）
        IF _eState = E_DL_SafetyDoorState.eFault THEN
            IF bDoorClosed AND bLockEngaged THEN
                _eState := E_DL_SafetyDoorState.eLocked; // 门锁全确认回闭锁态（重启抑制仍保持）/ Back to locked, inhibit retained
            ELSE
                _eState := E_DL_SafetyDoorState.eIdle;   // 否则回待机（Otherwise back to idle）
            END_IF
        END_IF
    END_IF
END_IF

// ============================================================================
// 段 3｜故障全局监视（优先级最高）
//      Global fault monitors (highest priority)
// ============================================================================
IF (NOT bDoorClosed) AND bLockEngaged THEN
    _bFaultLatch := TRUE;         // 门开+锁闭反馈同真：物理不可能组合，防篡改冲突锁存（Tamper conflict latch）
    _uErrorIdInt := 16#0003_0291; // 0003_0291 门锁不合理组合（防篡改冲突）【故障级】/ Impossible door-lock combination, fault level
    _eState := E_DL_SafetyDoorState.eFault;
ELSIF _fbTonUnlockTo.Q AND (_eState = E_DL_SafetyDoorState.eStopRequested) THEN
    _bFaultLatch := TRUE;         // 静止确认超时锁存（Standstill timeout latch）
    _uErrorIdInt := 16#0003_0290; // 0003_0290 静止确认超时（解锁链未达成）【故障级】/ Standstill confirmation timeout, fault level
    _eState := E_DL_SafetyDoorState.eFault;
ELSIF _fbTonRelockWin.Q AND _bRelockCheck THEN
    _bFaultLatch := TRUE;         // 再锁定超时锁存（Relock timeout latch）
    _uErrorIdInt := 16#0003_0292; // 0003_0292 再锁定超时【故障级】/ Relock timeout, fault level
    _eState := E_DL_SafetyDoorState.eFault;
    _bRelockCheck := FALSE;       // 确认窗计时终止（Confirm window terminated）
END_IF

// ============================================================================
// 段 4｜核心时序状态机（ENUM + CASE，含 ELSE 非法状态兜底）
//      Core sequence state machine (ENUM + CASE with ELSE fallback)
// ============================================================================
IF NOT _bFaultLatch THEN
    CASE _eState OF

        E_DL_SafetyDoorState.eIdle: // 待机态：门锁全确认，可受理解锁
            IF _bRestartInhibit THEN
                IF _fbTrigReset.Q THEN
                    _bRestartInhibit := FALSE;  // 复位沿解除重启抑制（Reset edge releases restart inhibit）
                END_IF
            ELSIF _bUnlockReq AND bDoorClosed AND bLockEngaged THEN
                _bPendUnlock := FALSE;          // 消费方法解锁请求（Consume method unlock）
                _eState := E_DL_SafetyDoorState.eStopRequested; // 进入解锁时序（Enter unlock sequence）
            ELSIF _bUnlockReq THEN
                _bPendUnlock := FALSE;          // 门锁未全确认的请求就地拒绝（Request rejected when door/lock not confirmed）
            END_IF

        E_DL_SafetyDoorState.eLocked: // 已闭锁态：再锁定确认中或重启抑制保持
            IF _bRelockCheck THEN
                IF bLockEngaged THEN
                    _bRelockCheck := FALSE;     // 窗内锁闭确认达成（Engagement confirmed inside window）
                END_IF                          // 超窗由段 3 全局监视接管（Window overrun handled by stage 3）
            ELSE
                IF _bRestartInhibit THEN
                    IF _fbTrigReset.Q THEN
                        _bRestartInhibit := FALSE; // 复位沿解除重启抑制（Reset edge releases inhibit）
                        _eState := E_DL_SafetyDoorState.eIdle; // 回待机（Back to idle）
                    END_IF
                ELSE
                    _eState := E_DL_SafetyDoorState.eIdle; // 无抑制直接回待机（No inhibit, back to idle）
                END_IF
            END_IF

        E_DL_SafetyDoorState.eStopRequested: // 已请求停机：等静止确认
            IF NOT bUseStandstillFb THEN
                _uInfoCode := 16#0003_0121;  // 0003_0121 run-down 计时器模式提示【信息级】（非零速实测）/ Run-down timer mode hint, info level
            END_IF
            IF bUseStandstillFb THEN
                _bStandstillOk := bStandstill; // 零速反馈模式（Zero-speed feedback mode）
            ELSE
                _bStandstillOk := _fbTonRunDown.Q; // run-down 计时模式（Run-down timer mode）
            END_IF
            IF _bStandstillOk THEN
                _eState := E_DL_SafetyDoorState.eStandstillConfirmed; // 静止确认达成（To standstill confirmed）
            END_IF

        E_DL_SafetyDoorState.eStandstillConfirmed: // 静止已确认：单拍过渡进解锁
            _eState := E_DL_SafetyDoorState.eUnlocked; // 进入解锁输出态（To unlocked state）

        E_DL_SafetyDoorState.eUnlocked: // 已解锁态：等待开门
            IF NOT bDoorClosed THEN
                uOpenCount := uOpenCount + 1;   // 开门审计累加（Open audit increment）
                _bRestartInhibit := TRUE;       // 开门事件置重启抑制（Open event arms restart inhibit）
                _eState := E_DL_SafetyDoorState.eOpened; // 转门开态（To opened state）
            END_IF

        E_DL_SafetyDoorState.eOpened: // 门已开启：等关门再锁定
            IF _bPendRelock OR bCmdRelock THEN
                _bPendRelock := FALSE;          // 消费方法再闭锁请求（Consume method relock）
            END_IF
            IF bDoorClosed THEN
                _bRelockCheck := TRUE;          // 关门沿启动再锁定确认窗（Door closed starts relock window）
                _eState := E_DL_SafetyDoorState.eLocked; // 转闭锁态（To locked state）
            END_IF

        E_DL_SafetyDoorState.eFault: // 故障锁存态：复位路径见段 2
            // 等待复位（Await reset）

        ELSE
            // 非法状态兜底：任何越界枚举值强制锁存故障（Illegal state fallback）
            _bFaultLatch := TRUE;           // 故障锁存（Fault latch）
            _uErrorIdInt := 16#0003_0293;   // 0003_0293 非法状态兜底【故障级】/ Illegal state, fault level
            _eState := E_DL_SafetyDoorState.eFault;
    END_CASE
END_IF

// ============================================================================
// 段 5｜输出推导 + 解锁电磁铁出口断言式硬约束
//      Output derivation + exit-assertion hard constraint of the unlock coil
// ============================================================================
// 解锁链硬约束：三条件不满足时解锁输出恒断（出口断言式写法）
// Hard constraint: the coil stays off unless all three conditions hold
IF _bStandstillOk AND bDoorClosed AND bLockEngaged AND (_eState = E_DL_SafetyDoorState.eUnlocked) AND (NOT _bFaultLatch) THEN
    bUnlockCoil := TRUE;              // 解锁电磁铁输出有效（Coil energized）
ELSE
    bUnlockCoil := FALSE;             // 出口断言恒断（Assertion: coil off）
END_IF
bStopRequest := (_eState = E_DL_SafetyDoorState.eStopRequested)
            OR (_eState = E_DL_SafetyDoorState.eStandstillConfirmed)
            OR (_eState = E_DL_SafetyDoorState.eUnlocked); // 停机请求随时序派生（Stop request follows the sequence）
IF _bFaultLatch THEN
    bStopRequest := FALSE;            // 故障态停机请求断（出口断言）/ Stop request forced off in fault (assertion)
END_IF

(*------------------------------------------------------------------------------
 * 方法: CmdRequestUnlock —— 请求解锁：发起停机请求并进入解锁时序。
 *      Method CmdRequestUnlock - starts the unlock sequence via stop request.
 *------------------------------------------------------------------------------*)

PROPERTY eState : E_DL_SafetyDoorState
eState := _eState;                // 返回内部状态（Return internal state）

(*------------------------------------------------------------------------------
 * 属性: bClosed（GET）—— 门已关闭反馈镜像。
 *      Property bClosed (GET) - door-closed feedback mirror.
 *------------------------------------------------------------------------------*)
PROPERTY bClosed : BOOL
bClosed := bDoorClosed;           // 反馈镜像（Feedback mirror）

(*------------------------------------------------------------------------------
 * 属性: bLocked（GET）—— 锁已闭锁反馈镜像。
 *      Property bLocked (GET) - lock-engaged feedback mirror.
 *------------------------------------------------------------------------------*)
PROPERTY bLocked : BOOL
bLocked := bLockEngaged;          // 反馈镜像（Feedback mirror）

(*------------------------------------------------------------------------------
 * 属性: bUnlockPermitted（GET）—— 允许解锁：无故障、无重启抑制且门锁全确认。
 *      Property bUnlockPermitted (GET) - unlock permitted derivation.
 *------------------------------------------------------------------------------*)
PROPERTY bUnlockPermitted : BOOL
bUnlockPermitted := (NOT _bFaultLatch) AND (NOT _bRestartInhibit)
                AND bDoorClosed AND bLockEngaged
                AND ((_eState = E_DL_SafetyDoorState.eIdle) OR (_eState = E_DL_SafetyDoorState.eLocked)); // 多条件派生式（Multi-condition derived form）

(*------------------------------------------------------------------------------
 * 属性: bOpened（GET）—— 门开启诊断镜像。
 *      Property bOpened (GET) - door-open diagnostic mirror.
 *------------------------------------------------------------------------------*)
PROPERTY bOpened : BOOL
bOpened := NOT bDoorClosed;       // 门开镜像（Door-open mirror）

(*------------------------------------------------------------------------------
 * 属性: bFault（GET）—— 故障锁存指示（信息级码不置本位，0.2 公约）。
 *      Property bFault (GET) - fault latch indicator, info codes excluded.
 *------------------------------------------------------------------------------*)
PROPERTY bFault : BOOL
bFault := _bFaultLatch OR (_eState = E_DL_SafetyDoorState.eFault); // 显式排除信息级派生式（Derived form excluding info codes）

(*------------------------------------------------------------------------------
 * 属性: uErrorId（GET）—— 末次故障码（故障级优先，无故障时透出本拍信息级
 *         码，0.2/0.15 公约）。
 *      Property uErrorId (GET) - last error code (fault priority, info shown otherwise).
 *------------------------------------------------------------------------------*)
PROPERTY uErrorId : UDINT
IF (_uErrorIdInt <> 0) OR (_eState = E_DL_SafetyDoorState.eFault) THEN
    uErrorId := _uErrorIdInt;     // 故障级码优先透出（Fault-level priority）
ELSE
    uErrorId := _uInfoCode;       // 无故障时透出本拍信息级码（Transient info code）
END_IF
END_FUNCTION_BLOCK
